(* IEC 61131-3 sources: daoli-st-library/DL_Process (part 53) *)

(* ---- FB_DL_StringCurrentMismatch.st ---- *)
(*
  FB_DL_StringCurrentMismatch  —  组串电流失配诊断与遮挡定位 / PV string current mismatch diagnostics and shading localisation
  分类 Category : DL_Process
  码位 Code     : 16#06_0_84
  版本 Version  : 1.0.0
  溯源 Source   : LGF Measurement 语义借鉴 · clean-room 实现，仅借分类/参数域/命名，未复制源码
  功能 Function : 1) 剔除无效/停机串后取中位基线（中位数抗单串遮挡污染，优于均值）；
                  2) 按失配率分级，失配率分母（基线）近零时自动切换为绝对差判据，防除零；
                  3) 输出最劣串物理串号（连续编址 1..16，越界钳位并置码）与失配掩码。
  边界 Boundary : ① 中位基线计算前剔除无效/停机串（电流 <= 0 或 NaN），有效样本 < 3 时不出诊断结论；
                  ② 失配率分母近零时改绝对差判据（防除零）；
                  ③ 遮挡定位输出按物理串号连续编址，越界下标钳位并置码；
                  ④ 结论态三行同向：基线值 → 最劣串号 → 失配标志。
  依赖 Depends  : None

  码表 Error codes（本件子码步进 16#10，避让邻件码位）:
    16#0002_0684 故障级：串数配置越界（nStringCount 不在 1..16）
    16#0002_0694 故障级：物理串号越界（枚举兜底路径，索引钳位后仍不可能命中）
    16#0002_06A4 信息级：有效样本不足 3 串，本轮不出诊断结论（不置 bError）
*)

TYPE E_DL_ScmPhase :
(
    eIdle    := 0,   // 空闲 / Idle
    eCollect := 10,  // 采样与剔除 / Sampling and rejection
    eDiagnose:= 20,  // 诊断计算 / Diagnostic computation
    eVerdict := 30,  // 结论输出 / Verdict output
    eFault   := 90   // 故障锁定 / Fault locked
);
END_TYPE

FUNCTION_BLOCK FB_DL_StringCurrentMismatch
VAR_INPUT
    bEnable       : BOOL;                         // 总使能，FALSE 回空闲 / Master enable
    bSample       : BOOL := TRUE;                 // 采样使能，TRUE 每拍纳入诊断 / Sampling enable
    bReset        : BOOL;                         // 复位，上升沿清故障 / Reset, clears fault
    nStringCount  : INT := 16;                    // 组串总数 [串]，域 1~16 / String count, 1..16
    afCurrentA    : ARRAY[1..16] OF REAL;         // 各串电流 [A]，域 > 0 为有效 / Per-string current [A]
    abStringValid : ARRAY[1..16] OF BOOL;         // 各串通讯/熔断有效标志 / Per-string valid flag
    fMismatchPct  : REAL := 10.0;                 // 失配率告警门限 [%]，域 0~100 / Mismatch rate alarm limit [%]
    fAbsFloorA    : REAL := 0.5;                  // 基线近零时的绝对差门限 [A]，域 > 0 / Absolute-difference limit [A]
    fBaselineEpsA : REAL := 0.1;                  // 基线近零判据容差 [A]，域 > 0 / Baseline near-zero tolerance [A]
    fMinSample    : INT := 3;                     // 最少有效样本数 [串]，常量 3 / Minimum valid sample count
END_VAR
VAR_OUTPUT
    fBaselineA    : REAL;                         // 中位基线电流 [A] / Median baseline current [A]
    nWorstIdx     : INT;                          // 最劣串物理串号 1..16，0 = 无 / Worst string number, 0 = none
    fWorstDevPct  : REAL;                         // 最劣串失配率 [%] / Worst string mismatch rate [%]
    fWorstDevA    : REAL;                         // 最劣串绝对偏差 [A] / Worst string absolute deviation [A]
    abMismatchMask : ARRAY[1..16] OF BOOL;        // 失配掩码 [开关]，索引 = 物理串号 / Mismatch mask per physical string
    nMismatchCount : INT;                         // 失配串数 [串] / Mismatched string count
    bMismatch     : BOOL;                         // 存在失配（保持型）/ Mismatch present, held
    bEnoughSample : BOOL;                         // 样本数满足结论条件 / Enough samples for a verdict
    bError        : BOOL;                         // 故障标志，与故障级码配对 / Fault flag paired with fault codes
    uErrorId      : UDINT;                        // 事件码，0 = 无事件 / Event code, 0 = none
    eStateOut     : E_DL_ScmPhase;                // 状态机当前态，段尾单点映射 / Phase mapped at tail
END_VAR
VAR
    _eState       : E_DL_ScmPhase := E_DL_ScmPhase.eIdle;  // 内部状态 / Internal state
    rtrReset      : R_TRIG;                       // 复位沿 / Reset edge
    nN            : INT;                          // 钳位后串数 [串] / Clamped string count
    nI            : INT;                          // 串循环下标 / String loop index
    nJ            : INT;                          // 排序内层下标 / Sort inner index
    nValid        : INT;                          // 有效串数 [串] / Valid string count
    nClampCode    : INT;                          // 下标钳位次数 [次] / Index clamping count
    afSort        : ARRAY[1..16] OF REAL;         // 有效电流排序缓存 [A] / Sorted valid currents [A]
    fTmp          : REAL;                         // 排序交换暂存 [A] / Sort swap buffer [A]
    fMedian       : REAL;                         // 中位基线暂存 [A] / Median baseline buffer [A]
    fDev          : REAL;                         // 单串偏差暂存 [A] / Single-string deviation [A]
    fRate         : REAL;                         // 单串失配率暂存 [%] / Single-string rate [%]
    fWorst        : REAL;                         // 最劣偏差累计 [A] / Worst deviation accumulator [A]
    bNearZero     : BOOL;                         // 基线近零标志 / Baseline near-zero flag
    uFault        : UDINT;                        // 锁存故障码 / Latched fault code
    uInfo         : UDINT;                        // 信息级码 / Information code
END_VAR
VAR CONSTANT
    DL_SCM_STRMAX : INT := 16;                    // 组串数组上界 [串] / String array upper bound
    DL_SCM_PCTMAX : REAL := 100.0;                // 失配率上限 [%] / Mismatch rate ceiling [%]
END_VAR

(* === 段 0 · 实例刷新（无条件周期调用）=== *)
rtrReset(CLK := bReset);                          // 每拍刷新复位沿

(* === 段 1 · 组态与索引闸 === *)
nN := nStringCount;                               // 串数取用前钳位
IF nN < 1 THEN
    nN := 1;                                      // 下限钳位
END_IF
IF nN > DL_SCM_STRMAX THEN
    nN := DL_SCM_STRMAX;                          // 上限钳位
END_IF
IF (nStringCount < 1) OR (nStringCount > DL_SCM_STRMAX) THEN
    uFault := 16#0002_0684;                       // 故障级：串数配置越界
END_IF
IF rtrReset.Q THEN
    uFault := 16#0000;                            // 复位沿清锁存
    bMismatch := FALSE;                           // 失配标志同步复位
    nWorstIdx := 0;                               // 最劣串号复位
END_IF

(* === 段 2 · 主状态机（ENUM + CASE，含 ELSE 兜底）=== *)
CASE _eState OF
E_DL_ScmPhase.eIdle :
    bEnoughSample := FALSE;                       // 空闲无结论
    uInfo := 16#0000;                             // 信息码清零
    IF uFault = 16#0002_0684 THEN
        _eState := E_DL_ScmPhase.eFault;          // 组态故障优先
    ELSIF bEnable AND bSample THEN
        _eState := E_DL_ScmPhase.eCollect;        // 本拍进入采样相
    END_IF

E_DL_ScmPhase.eCollect :
    nValid := 0;                                  // 有效串计数清零
    nClampCode := 0;                              // 钳位计数清零
    FOR nI := 1 TO DL_SCM_STRMAX DO
        IF nI <= nN THEN
            IF abStringValid[nI]
               AND (afCurrentA[nI] = afCurrentA[nI])              // NaN 自反判据
               AND (ABS(afCurrentA[nI]) < 1.0E30)                 // Inf 上限兜底
               AND (afCurrentA[nI] > 0.0) THEN                    // 停机串（<= 0）剔除
                nValid := nValid + 1;                             // 有效样本计数
                afSort[nValid] := afCurrentA[nI];                 // 收入排序缓存，nValid 已受 DL_SCM_STRMAX 约束
            END_IF
        END_IF
    END_FOR
    IF fMinSample < 3 THEN
        fMinSample := 3;                          // 最小样本数下限钳位（域 >= 3，防组态放宽到误判）
    END_IF
    bEnoughSample := (nValid >= fMinSample);      // 样本不足不出结论
    IF bEnoughSample THEN
        _eState := E_DL_ScmPhase.eDiagnose;       // 转诊断相
    ELSE
        uInfo := 16#0002_06A4;                    // 信息级：样本不足
        _eState := E_DL_ScmPhase.eVerdict;        // 仍走结论相，但结论为空
    END_IF

E_DL_ScmPhase.eDiagnose :
    FOR nI := 1 TO (nValid - 1) DO                // 插入排序求中位数
        FOR nJ := nI + 1 TO nValid DO
            IF afSort[nJ] < afSort[nI] THEN
                fTmp := afSort[nI];               // 交换暂存
                afSort[nI] := afSort[nJ];
                afSort[nJ] := fTmp;
            END_IF
        END_FOR
    END_FOR
    IF (nValid MOD 2) = 1 THEN
        fMedian := afSort[(nValid + 1) / 2];      // 奇数：取正中样本，下标受 nValid 约束
    ELSE
        fMedian := (afSort[nValid / 2] + afSort[(nValid / 2) + 1]) * 0.5;   // 偶数：取中两样本均值
    END_IF
    fBaselineA := fMedian;                        // 基线输出
    bNearZero := (ABS(fMedian) <= fBaselineEpsA); // 基线近零判据（防除零前置）
    nWorstIdx := 0;                               // 最劣串号先清零
    fWorst := -1.0;                               // 最劣偏差累计初值（负值确保首次必更新）
    fWorstDevPct := 0.0;                          // 最劣失配率初值
    fWorstDevA := 0.0;                            // 最劣绝对偏差初值
    nMismatchCount := 0;                          // 失配串计数清零
    FOR nI := 1 TO DL_SCM_STRMAX DO
        abMismatchMask[nI] := FALSE;              // 掩码逐串先清零
        IF nI <= nN THEN
            IF abStringValid[nI] AND (afCurrentA[nI] = afCurrentA[nI]) AND (afCurrentA[nI] > 0.0) THEN
                fDev := fMedian - afCurrentA[nI];                 // 偏差 = 基线 − 实测（正 = 偏低）
                IF bNearZero THEN
                    fRate := ABS(fDev);                               // 基线近零：改绝对差判据
                ELSE
                    fRate := ABS(fDev) / ABS(fMedian) * DL_SCM_PCTMAX;   // 分母已判非零
                END_IF
                IF fRate > DL_SCM_PCTMAX THEN
                    fRate := DL_SCM_PCTMAX;                       // 失配率饱和，防超界显示
                END_IF
                IF (bNearZero AND (ABS(fDev) > fAbsFloorA))
                   OR ((NOT bNearZero) AND (fRate >= fMismatchPct)) THEN
                    abMismatchMask[nI] := TRUE;                   // 该串判失配
                    nMismatchCount := nMismatchCount + 1;         // 失配计数累加
                END_IF
                IF fDev > fWorst THEN
                    fWorst := fDev;                               // 记录最劣偏差
                    IF (nI >= 1) AND (nI <= DL_SCM_STRMAX) THEN
                        nWorstIdx := nI;                          // 物理串号连续编址
                    ELSE
                        nWorstIdx := 0;                           // 越界下标钳位为 0
                        nClampCode := nClampCode + 1;             // 记录钳位事件
                    END_IF
                    fWorstDevPct := fRate;                        // 最劣串失配率
                    fWorstDevA := ABS(fDev);                      // 最劣串绝对偏差
                END_IF
            END_IF
        END_IF
    END_FOR
    bMismatch := (nMismatchCount > 0);            // 置位型结论：存在失配（段尾不清零）
    IF nClampCode > 0 THEN
        uFault := 16#0002_0694;                   // 故障级：物理串号越界已钳位
    END_IF
    _eState := E_DL_ScmPhase.eVerdict;            // 转结论相

E_DL_ScmPhase.eVerdict :
    IF NOT bEnoughSample THEN
        nWorstIdx := 0;                           // 样本不足：不给定位结论
        nMismatchCount := 0;                      // 失配计数归 0
        fWorstDevPct := 0.0;                      // 失配率归 0，避免误导
    END_IF
    IF (NOT bEnable) OR rtrReset.Q THEN
        _eState := E_DL_ScmPhase.eIdle;           // 失能/复位回空闲
    ELSIF bSample THEN
        _eState := E_DL_ScmPhase.eCollect;        // 连续采样：下一拍重新采集
    END_IF

E_DL_ScmPhase.eFault :
    bEnoughSample := FALSE;                       // 故障态不出结论
    nWorstIdx := 0;                               // 最劣串号 0
    IF uFault = 16#0000 THEN
        _eState := E_DL_ScmPhase.eIdle;           // 解锁后回空闲
    END_IF

ELSE
    _eState := E_DL_ScmPhase.eFault;              // 非法状态拦截
    uFault := 16#0002_0694;                       // 故障级：相 ID 越界（枚举兜底路径）
END_CASE

(* === 段 3 · 输出映射（三行同向：基线 → 最劣串号 → 失配标志）=== *)
IF NOT bEnoughSample THEN
    fBaselineA := fMedian;                        // 基线仍输出（诊断可读）
    bMismatch := nMismatchCount > 0;               // 失配标志与计数严格同源
END_IF
IF NOT bEnable THEN
    bMismatch := FALSE;                           // 失能强制清失配结论
    nWorstIdx := 0;                               // 最劣串号归 0
END_IF
bError := (uFault <> 16#0000);                    // 故障标志仅由故障级码置位（R45 配对）
IF bError THEN
    uErrorId := uFault;                           // 故障级优先上报
ELSE
    uErrorId := uInfo;                            // 否则上报信息级码
END_IF
eStateOut := _eState;                             // 输出枚举段尾单点映射（N2 规则）
END_FUNCTION_BLOCK

(* ---- FB_DL_StringElImageMap.st ---- *)
(*
  ==================================================================
  组件名 Component  : FB_DL_StringElImageMap
  分类   Category   : DL_Process
  版本   Version    : 1.0.1
  功能   Purpose    : EL 图像缺陷坐标归档与批次比对。逐条接收缺陷报告（坐标、面积、
                      类型），回钳后写入环窗归档（最新 64 条），并按批号累计本批
                      缺陷数、面积和 / 最大值 / 类型掩码；批号变化沿把当前批统计
                      转入「上批」快照并清零当前批，随后给出与上批的比对结论
                      （缺陷数与最大面积双向带容差比较）。
  溯源   Origin     : 缺陷坐标归档与批次间对比为通用视觉质量统计语义；本件为
                      clean-room 实现，仅借鉴来源分类与参数域组织（来源标签
                      roadmap-p2-elimage），道莅原创设计，未复制任何闭源代码行。
  平台   Platform   : 纯 IEC 61131-3（ARRAY / WORD / SHL / R_TRIG，无私有库）
  作者   Author     : 道莅代码库 · PLC 编程专家（R55）
  ------------------------------------------------------------------
  边界 Boundary     :
                      一 本件只做归档与统计比对，不做缺陷判定、不存图像（属主边界）；
                      二 坐标越出视野范围不归档，但计入越界计数并置信息级成因；
                      三 非有限坐标或面积不归档、不计数，出口数值保持上拍值；
                      四 环窗游标一律经回钳 1..64，写入顺序为「先算槽位、后写入」；
                      五 无全局变量、无外部变量声明、无物理地址寻址。
  输出契约 Output contract:
                      wTypeMask 位 i-1 对应缺陷类型 i（类型 1 得 bit0，类型 8 得 bit7）；
                      bComparePass 仅在无参照批（上批缺陷数为零）时恒为真，
                      有参照批时按「缺陷数」与「最大面积」双向带容差比较；
                      eCause 故障级成因与 bError 配对（R45），信息级永不置 bError。
  修订记录 Revision  :
    2026-11-20  v1.0.0  R55 首版（批 3 · 序号 12）
    2026-11-20  v1.0.1  R56 返修（7.4）：段 2 复位作用域补清 fLastXmm / fLastYmm /
                        fLastSizeMm2 / nLastType 四个最近缺陷出口，并补
                        _stCur.uBatchId 批号重同步，防复位后首条新批报告误判入旧批窗口。
  ==================================================================
*)

TYPE ST_DL_ElBatchStat :
STRUCT
    uBatchId  : UDINT := 0;      // 批号 [-] / batch identifier
    nCount    : INT := 0;        // 缺陷条数 [条] / defect count [piece]
    fSumSize  : REAL := 0.0;     // 面积累计 [平方毫米] / accumulated area [square millimetre]
    fMaxSize  : REAL := 0.0;     // 面积最大值 [平方毫米] / maximum area [square millimetre]
    wTypeMask : WORD := 16#0000; // 类型掩码 [-] / type mask
END_STRUCT
END_TYPE

TYPE E_DL_SeiCause :
(
    eNone       := 0,   // 无成因 / no cause
    eCfgIllegal := 1,   // 组态非法：视野范围或容差越域（故障级，与 bError 配对）/ illegal config, field bounds or tolerance out of domain
    eOutField   := 2,   // 缺陷坐标越出视野，未归档（信息级）/ the defect coordinate is outside the field and was not archived, informational
    eInputBad   := 3,   // 坐标或面积非有限，未归档（信息级）/ non-finite coordinate or area, not archived, informational
    eTypeBad    := 4    // 缺陷类型越域已回钳（信息级）/ the defect type was clamped, informational
);
END_TYPE

FUNCTION_BLOCK FB_DL_StringElImageMap
VAR_INPUT
    bEnable       : BOOL := TRUE;            // 使能，失能时不接收缺陷报告 [-] / enable, defect reports are not accepted when disabled
    bReset        : BOOL := FALSE;          // 复位上升沿清故障锁存与全部统计 [-] / reset rising edge clears the fault latch and all statistics
    bDefectValid  : BOOL := FALSE;           // 缺陷报告脉冲，上升沿归档一次 [-] / defect report pulse, archived once on the rising edge
    fPosXmm       : REAL := 0.0;             // 缺陷中心横坐标 [毫米] / defect centre abscissa [millimetre]
    fPosYmm       : REAL := 0.0;             // 缺陷中心纵坐标 [毫米] / defect centre ordinate [millimetre]
    fSizeMm2      : REAL := 0.0;             // 缺陷面积 [平方毫米] / defect area [square millimetre]
    nDefectType   : INT := 1;                // 缺陷类型 [类型号]，域 1..8 / defect type [type number], domain 1 to 8
    uBatchId      : UDINT := 0;              // 当前批号 [-] / current batch identifier
    fFieldXmm     : REAL := 1000.0;          // 视野横向范围 [毫米]，域 大于零 / field width [millimetre], domain above zero
    fFieldYmm     : REAL := 1000.0;          // 视野纵向范围 [毫米]，域 大于零 / field height [millimetre], domain above zero
    fTolPct       : REAL := 10.0;            // 批次比对容差 [百分比]，域 大于零 / batch comparison tolerance [percent], domain above zero
END_VAR
VAR_OUTPUT
    fLastXmm      : REAL := 0.0;             // 最近归档缺陷横坐标 [毫米] / abscissa of the last archived defect [millimetre]
    fLastYmm      : REAL := 0.0;             // 最近归档缺陷纵坐标 [毫米] / ordinate of the last archived defect [millimetre]
    fLastSizeMm2  : REAL := 0.0;             // 最近归档缺陷面积 [平方毫米] / area of the last archived defect [square millimetre]
    nLastType     : INT := 0;                // 最近归档缺陷类型 [类型号] / type of the last archived defect [type number]
    uArchiveCnt   : UDINT := 0;              // 累计归档缺陷数 [条] / total archived defects [piece]
    nBufCount     : INT := 0;                // 环窗当前条数 [条] / ring buffer occupancy [piece]
    nCurCount     : INT := 0;                // 当前批缺陷条数 [条] / current batch defect count [piece]
    fCurMaxMm2    : REAL := 0.0;             // 当前批最大缺陷面积 [平方毫米] / current batch maximum area [square millimetre]
    fCurMeanMm2   : REAL := 0.0;             // 当前批平均缺陷面积 [平方毫米] / current batch mean area [square millimetre]
    nPrevCount    : INT := 0;                // 上批缺陷条数 [条] / previous batch defect count [piece]
    fPrevMaxMm2   : REAL := 0.0;             // 上批最大缺陷面积 [平方毫米] / previous batch maximum area [square millimetre]
    fDeltaMaxPct  : REAL := 0.0;             // 最大面积相对变化 [百分比] / relative change of the maximum area [percent]
    bComparePass  : BOOL := FALSE;           // 批次比对通过 [-] / batch comparison passed
    wTypeMask     : WORD := 16#0000;         // 当前批缺陷类型掩码 [-] / current batch defect type mask
    nOutFieldCnt  : INT := 0;                // 越界缺陷计数（饱和到上限）[条] / out of field defect count, saturated [piece]
    eCause        : E_DL_SeiCause := E_DL_SeiCause.eNone; // 成因出口 [枚举] / cause outlet [enum]
    bError        : BOOL := FALSE;           // 故障锁存标志 [-] / fault latch flag
END_VAR
VAR
    rtDefect      : R_TRIG;                  // 缺陷报告沿检测，段 0 无条件刷新 / defect report edge detector, refreshed unconditionally in segment zero
    rtReset       : R_TRIG;                  // 复位沿检测，段 0 无条件刷新 / reset edge detector, refreshed unconditionally in segment zero
    _stCur        : ST_DL_ElBatchStat;       // 当前批统计 / current batch statistics
    _stPrev       : ST_DL_ElBatchStat;       // 上批统计快照 / previous batch statistics snapshot
    _eCause       : E_DL_SeiCause := E_DL_SeiCause.eNone;  // 信息级成因，每拍重算 / informational cause, recomputed every scan
    _eFaultCause  : E_DL_SeiCause := E_DL_SeiCause.eNone;  // 故障级成因，锁存至复位沿 / fault cause, latched until the reset edge
    _bFault       : BOOL := FALSE;           // 故障锁存位 [-] / fault latch bit
    _bInit        : BOOL := FALSE;           // 首扫初始化完成标志（R310）/ first scan initialisation flag
    _bCfgBad      : BOOL := FALSE;           // 组态非法判定 [-] / illegal configuration verdict
    _bInOk        : BOOL := FALSE;           // 本拍缺陷数据有限 [-] / this scan defect data finite
    _bInField     : BOOL := FALSE;           // 坐标在视野内 [-] / the coordinate is inside the field
    _bTypeClamped : BOOL := FALSE;           // 类型号被回钳 [-] / the type number was clamped
    _bBatchRoll   : BOOL := FALSE;           // 本拍发生批号变化 [-] / the batch identifier changed this scan
    _nTypeUse     : INT := 1;                // 钳定后的缺陷类型号 [类型号] / clamped defect type number
    _nIdx         : INT := 1;                // 环窗写入槽位（1 起，回钳 1..64）[槽号] / ring write slot, one-based, clamped one through sixty four
    _wTypeBit     : WORD := 16#0001;         // 类型位掩码，先移位后置位（R327）/ type bit mask, shift before setting
    _wMask        : WORD := 16#0000;         // 类型掩码工作字 / type mask working word
    _fMean        : REAL := 0.0;             // 均值工作值 [平方毫米] / mean working value [square millimetre]
    _fDeltaPct    : REAL := 0.0;             // 相对变化工作值 [百分比] / relative change working value [percent]
    _fPrevMaxB    : REAL := 0.0;             // 上批最大面积基线，用于除零闸 [平方毫米] / previous maximum baseline against division by zero [square millimetre]
    _fPrevCntB    : REAL := 0.0;             // 上批条数基线，用于除零闸 [条] / previous count baseline against division by zero [piece]
    _fCurMaxB     : REAL := 0.0;             // 当前批最大面积暂存 [平方毫米] / current maximum area held in a local [square millimetre]
    _fCurCntB     : REAL := 0.0;             // 当前批条数暂存 [条] / current count held in a local [piece]
    _afX          : ARRAY[1..64] OF REAL := [64(0.0)]; // 环窗横坐标归档 [毫米] / ring archive of abscissae [millimetre]
    _afY          : ARRAY[1..64] OF REAL := [64(0.0)]; // 环窗纵坐标归档 [毫米] / ring archive of ordinates [millimetre]
    _afSz         : ARRAY[1..64] OF REAL := [64(0.0)]; // 环窗面积归档 [平方毫米] / ring archive of areas [square millimetre]
    _anType       : ARRAY[1..64] OF INT := [64(0)];    // 环窗类型归档 [类型号] / ring archive of type numbers [type number]
END_VAR
VAR CONSTANT
    DL_SEI_BUF_MAX   : INT := 64;            // 环窗容量与槽位回钳上界 [条] / ring capacity and slot clamp upper bound
    DL_SEI_TYPE_MIN  : INT := 1;             // 缺陷类型下限 [类型号] / defect type floor [type number]
    DL_SEI_TYPE_MAX  : INT := 8;             // 缺陷类型上限（与掩码位宽一致）[类型号] / defect type ceiling matching the mask width [type number]
    DL_SEI_COUNT_MAX : INT := 30000;         // 单批缺陷条数上限，防溢出 [条] / per batch defect count ceiling against overflow [piece]
    DL_SEI_AREA_MAX  : REAL := 1.0E6;        // 缺陷面积量级上限 [平方毫米] / defect area magnitude ceiling [square millimetre]
    DL_SEI_TOL_MAX   : REAL := 500.0;        // 比对容差上限 [百分比] / comparison tolerance ceiling [percent]
    DL_SEI_MASK_NONE : WORD := 16#0000;      // 空掩码常量 [-] / empty mask constant
    DL_SEI_MASK_ONE  : WORD := 16#0001;      // 单位位常量 [-] / single bit constant
END_VAR

// 段 0｜沿检测无条件周期刷新（禁入分支）/ segment 0, unconditional refresh of the edge detectors, never inside a branch
rtDefect(CLK := bDefectValid); // 缺陷报告沿无条件刷新 / unconditional refresh of the defect edge
rtReset(CLK := bReset); // 复位沿无条件刷新 / unconditional refresh of the reset edge

// 段 1｜首扫初始化（R310）：统计与环窗从确定起点开始 / segment 1, first scan initialisation
IF NOT _bInit THEN // 首扫一拍 / the very first scan
    _bInit := TRUE; // 置首扫完成标志 / raise the first scan flag
    _bFault := FALSE; // 故障锁存清零 / clear the fault latch
    _eCause := E_DL_SeiCause.eNone; // 信息级成因清零 / clear the informational cause
    _eFaultCause := E_DL_SeiCause.eNone; // 故障级成因清零 / clear the fault cause
    _stCur.uBatchId := uBatchId; // 当前批号初始化 / initialise the current batch identifier
    _stPrev.uBatchId := 0; // 上批号清零 / clear the previous batch identifier
    _nIdx := 1; // 环窗槽位归位 / park the ring slot at one
END_IF

// 段 2｜复位沿作用域：清锁存 / 清统计 / 清环窗游标（归档数组保留，不作判据）/ segment 2, reset edge scope
IF rtReset.Q THEN // 复位沿 / reset edge
    _bFault := FALSE; // 作用域一：清故障锁存 / scope one, clear the fault latch
    _eFaultCause := E_DL_SeiCause.eNone; // 作用域一：清故障级成因 / scope one, clear the fault cause
    _stCur.nCount := 0; // 作用域二：清当前批条数 / scope two, clear the current batch count
    _stCur.fSumSize := 0.0; // 作用域二：清面积累计 / scope two, clear the accumulated area
    _stCur.fMaxSize := 0.0; // 作用域二：清面积最大值 / scope two, clear the maximum area
    _stCur.wTypeMask := DL_SEI_MASK_NONE; // 作用域二：清类型掩码 / scope two, clear the type mask
    _stPrev.nCount := 0; // 作用域二：清上批条数 / scope two, clear the previous count
    _stPrev.fSumSize := 0.0; // 作用域二：清上批面积累计 / scope two, clear the previous accumulated area
    _stPrev.fMaxSize := 0.0; // 作用域二：清上批最大面积 / scope two, clear the previous maximum area
    _stPrev.wTypeMask := DL_SEI_MASK_NONE; // 作用域二：清上批类型掩码 / scope two, clear the previous type mask
    fLastXmm := 0.0; // 作用域二：清最近横坐标出口（R56 返修补齐）/ scope two, clear the last abscissa outlet
    fLastYmm := 0.0; // 作用域二：清最近纵坐标出口（R56 返修补齐）/ scope two, clear the last ordinate outlet
    fLastSizeMm2 := 0.0; // 作用域二：清最近面积出口（R56 返修补齐）/ scope two, clear the last area outlet
    nLastType := 0; // 作用域二：清最近类型出口（R56 返修补齐）/ scope two, clear the last type outlet
    _stCur.uBatchId := uBatchId; // 作用域二：当前批号重同步，防复位后首条新批报告误判入旧批窗口（R56 返修补齐）/ scope two, resync the current batch identifier so the first report after a reset is not judged against a stale batch window
    _nIdx := 1; // 作用域三：清环窗槽位 / scope three, clear the ring slot cursor
    nBufCount := 0; // 作用域三：清环窗占用 / scope three, clear the ring occupancy
    uArchiveCnt := 0; // 作用域三：清累计归档数 / scope three, clear the total archived count
    nOutFieldCnt := 0; // 作用域三：清越界计数 / scope three, clear the out of field count
END_IF

// 段 3｜组态域闸（R151 全覆盖）：视野范围与比对容差 / segment 3, configuration domain gate over the field bounds and the tolerance
_bCfgBad := FALSE; // 组态非法预置假 / preset the illegal configuration verdict to false
IF (fFieldXmm <= 0.0) OR (fFieldXmm <> fFieldXmm) OR (fFieldXmm > DL_SEI_AREA_MAX) THEN // 横向视野越域 / field width out of domain
    _bCfgBad := TRUE; // 判非法 / mark illegal
END_IF
IF (fFieldYmm <= 0.0) OR (fFieldYmm <> fFieldYmm) OR (fFieldYmm > DL_SEI_AREA_MAX) THEN // 纵向视野越域 / field height out of domain
    _bCfgBad := TRUE; // 判非法 / mark illegal
END_IF
IF (fTolPct <= 0.0) OR (fTolPct > DL_SEI_TOL_MAX) OR (fTolPct <> fTolPct) THEN // 容量越域 / tolerance out of domain
    _bCfgBad := TRUE; // 判非法 / mark illegal
END_IF
IF _bCfgBad AND (NOT _bFault) THEN // 组态非法且未锁存 / illegal configuration and not yet latched
    _bFault := TRUE; // 置故障锁存 / raise the fault latch
    _eFaultCause := E_DL_SeiCause.eCfgIllegal; // 故障级成因 (R45 配对 bError) / fault grade cause paired with bError
END_IF

// 段 4｜批号变化：当前批统计转入上批快照，当前批清零 / segment 4, batch change moves the current statistics into the previous snapshot
_bBatchRoll := (uBatchId <> _stCur.uBatchId); // 批号变化判据 / batch change criterion
IF _bBatchRoll THEN // 批号变化 / the batch identifier changed
    _stPrev.uBatchId := _stCur.uBatchId; // 上批号继承 / the previous identifier inherits
    _stPrev.nCount := _stCur.nCount; // 上批条数快照 / snapshot the previous count
    _stPrev.fSumSize := _stCur.fSumSize; // 上批面积累计快照 / snapshot the previous accumulated area
    _stPrev.fMaxSize := _stCur.fMaxSize; // 上批最大面积快照 / snapshot the previous maximum area
    _stPrev.wTypeMask := _stCur.wTypeMask; // 上批类型掩码快照 / snapshot the previous type mask
    _stCur.uBatchId := uBatchId; // 当前批号推进 / advance the current identifier
    _stCur.nCount := 0; // 当前批条数清零 / clear the current count
    _stCur.fSumSize := 0.0; // 当前批面积累计清零 / clear the current accumulated area
    _stCur.fMaxSize := 0.0; // 当前批最大面积清零 / clear the current maximum area
    _stCur.wTypeMask := DL_SEI_MASK_NONE; // 当前批类型掩码清零 / clear the current type mask
END_IF

// 段 5｜缺陷归档：有限性闸 → 视野闸 → 类型回钳 → 环窗写入 → 统计累加 / segment 5, defect archiving chain
_eCause := E_DL_SeiCause.eNone; // 信息级成因每拍重算 / the informational cause is recomputed every scan
_bTypeClamped := FALSE; // 类型回钳标志预置假 / preset the type clamp flag to false
IF rtDefect.Q AND bEnable AND (NOT _bFault) THEN // 缺陷报告沿且使能无故障 / defect edge while enabled and unfaulted
    _bInOk := (fPosXmm = fPosXmm) AND ((fPosXmm - fPosXmm) = (fPosXmm - fPosXmm)) AND (fPosYmm = fPosYmm) AND ((fPosYmm - fPosYmm) = (fPosYmm - fPosYmm)) AND (fSizeMm2 = fSizeMm2) AND ((fSizeMm2 - fSizeMm2) = (fSizeMm2 - fSizeMm2)); // 坐标与面积有限性闸 / finiteness gate on coordinates and area
    _bInField := _bInOk AND (fPosXmm >= 0.0) AND (fPosXmm <= fFieldXmm) AND (fPosYmm >= 0.0) AND (fPosYmm <= fFieldYmm) AND (fSizeMm2 >= 0.0) AND (fSizeMm2 <= DL_SEI_AREA_MAX); // 视野与面积域闸 / field and area domain gate
    _nTypeUse := nDefectType; // 类型号直通 / the type number passes through
    IF _nTypeUse < DL_SEI_TYPE_MIN THEN // 下越界 / below the lower bound
        _nTypeUse := DL_SEI_TYPE_MIN; // 回钳到 1 / clamp to one
        _bTypeClamped := TRUE; // 置回钳标志 / raise the clamp flag
    ELSIF _nTypeUse > DL_SEI_TYPE_MAX THEN // 上越界 / above the upper bound
        _nTypeUse := DL_SEI_TYPE_MAX; // 回钳到 8 / clamp to eight
        _bTypeClamped := TRUE; // 置回钳标志 / raise the clamp flag
    END_IF
    IF NOT _bInOk THEN // 数据非有限 / data non-finite
        _eCause := E_DL_SeiCause.eInputBad; // 信息级成因：未归档 / informational cause, not archived
    ELSIF NOT _bInField THEN // 坐标或面积越域 / coordinate or area out of domain
        _eCause := E_DL_SeiCause.eOutField; // 信息级成因：越界未归档 / informational cause, out of field
        IF nOutFieldCnt < DL_SEI_COUNT_MAX THEN // 未达计数上限 / below the count ceiling
            nOutFieldCnt := nOutFieldCnt + 1; // 越界计数递增 / increment the out of field count
        END_IF
    ELSE
        // 段 5.1｜环窗写入：先算槽位再写入，槽位经回钳 1..64 / segment 5.1, ring write with the slot clamped one through sixty four
        _nIdx := _nIdx + 1; // 槽位前移 / advance the slot
        IF _nIdx > DL_SEI_BUF_MAX THEN // 越过上界 / past the upper bound
            _nIdx := 1; // 回钳到一号槽 / clamp back to slot one
        END_IF
        _afX[_nIdx] := fPosXmm; // 横坐标归档 / archive the abscissa
        _afY[_nIdx] := fPosYmm; // 纵坐标归档 / archive the ordinate
        _afSz[_nIdx] := fSizeMm2; // 面积归档 / archive the area
        _anType[_nIdx] := _nTypeUse; // 类型归档 / archive the type
        IF nBufCount < DL_SEI_BUF_MAX THEN // 环窗未满 / the ring is not yet full
            nBufCount := nBufCount + 1; // 占用递增 / increment the occupancy
        END_IF
        IF uArchiveCnt < 2000000000 THEN // 累计计数未达保护上限（常量在 DINT 可表范围内）/ the total count is below the guard ceiling, the constant fits in DINT
            uArchiveCnt := uArchiveCnt + 1; // 累计归档数递增 / increment the total archived count
        END_IF
        fLastXmm := fPosXmm; // 最近横坐标出口 / last abscissa outlet
        fLastYmm := fPosYmm; // 最近纵坐标出口 / last ordinate outlet
        fLastSizeMm2 := fSizeMm2; // 最近面积出口 / last area outlet
        nLastType := _nTypeUse; // 最近类型出口 / last type outlet
        // 段 5.2｜当前批统计累加 / segment 5.2, accumulate the current batch statistics
        IF _stCur.nCount < DL_SEI_COUNT_MAX THEN // 未达条数上限 / below the count ceiling
            _stCur.nCount := _stCur.nCount + 1; // 条数递增 / increment the count
        END_IF
        _stCur.fSumSize := _stCur.fSumSize + fSizeMm2; // 面积累计 / accumulate the area
        IF fSizeMm2 > _stCur.fMaxSize THEN // 面积最大值刷新 / refresh the maximum area
            _stCur.fMaxSize := fSizeMm2; // 更新最大值 / update the maximum
        END_IF
        _wTypeBit := SHL(DL_SEI_MASK_ONE, _nTypeUse - 1); // 类型位掩码，位移量 0..7 由类型回钳证明 / type bit mask, the shift zero through seven is proven by the type clamp
        _stCur.wTypeMask := _stCur.wTypeMask OR _wTypeBit; // 类型掩码置位 / set the type bit
        IF _bTypeClamped THEN // 类型被回钳 / the type was clamped
            _eCause := E_DL_SeiCause.eTypeBad; // 信息级成因 / informational cause
        END_IF
    END_IF
END_IF

// 段 6｜批次比对：双向带容差比较，参照批缺陷数为零时判通过 / segment 6, batch comparison with a two sided tolerance
_fCurMaxB := _stCur.fMaxSize; // 当前批最大面积 / the current maximum area
_fCurCntB := INT_TO_REAL(_stCur.nCount); // 当前批条数实数化 / the current count as a real
_fPrevMaxB := _stPrev.fMaxSize; // 上批最大面积 / the previous maximum area
_fPrevCntB := INT_TO_REAL(_stPrev.nCount); // 上批条数实数化 / the previous count as a real
IF (_fPrevMaxB > 0.0) THEN // 有参照批 / a reference batch exists
    _fDeltaPct := (_fCurMaxB - _fPrevMaxB) / _fPrevMaxB * 100.0; // 最大面积相对变化，除子已证大于零 / relative change of the maximum area, divisor proven positive
    bComparePass := (_fCurMaxB <= _fPrevMaxB * (1.0 + fTolPct / 100.0)) AND (_fPrevCntB <= 0.0 OR (_fCurCntB <= _fPrevCntB * (1.0 + fTolPct / 100.0))); // 数与面积双向比较，条数基线为零时只比面积 / the count and area are both compared, with a zero count baseline only the area is compared
ELSE // 无参照批 / no reference batch
    _fDeltaPct := 0.0; // 相对变化记零 / the relative change is zeroed
    bComparePass := TRUE; // 无参照按通过处理（不误判不合格）/ no reference passes so nothing is falsely rejected
END_IF

// 段 7｜统一出口 / segment 7, unified outlet
nCurCount := _stCur.nCount; // 当前批条数出口 / current count outlet
fCurMaxMm2 := _stCur.fMaxSize; // 当前批最大面积出口 / current maximum area outlet
_fMean := 0.0; // 均值预置零 / preset the mean to zero
IF _stCur.nCount > 0 THEN // 有条数才可算均值 / the mean needs at least one piece
    _fMean := _stCur.fSumSize / INT_TO_REAL(_stCur.nCount); // 均值，除子已证大于零 / mean, divisor proven positive
END_IF
fCurMeanMm2 := _fMean; // 当前批均值出口 / current mean outlet
nPrevCount := _stPrev.nCount; // 上批条数出口 / previous count outlet
fPrevMaxMm2 := _stPrev.fMaxSize; // 上批最大面积出口 / previous maximum area outlet
fDeltaMaxPct := _fDeltaPct; // 相对变化出口 / relative change outlet
wTypeMask := _stCur.wTypeMask; // 类型掩码出口 / type mask outlet
IF _bFault THEN // 故障锁存优先 / the fault latch takes priority
    eCause := _eFaultCause; // 故障级成因锁存回放 / the fault cause is replayed from the latch
ELSE
    eCause := _eCause; // 信息级成因直映 / the informational cause is mapped directly
END_IF
bError := _bFault; // 故障标志与锁存位同源 / the fault flag shares the latch source
END_FUNCTION_BLOCK

(* ---- FB_DL_StringerTrend.st ---- *)
(*
  FB_DL_StringerTrend  —  串焊机多通道焊接温度曲线在线监视 / Stringer multi-channel soldering temperature monitor
  分类 Category : DL_Process
  码位 Code     : 16#06_0_8E
  版本 Version  : 1.0.0
  溯源 Source   : LGF Measurement 语义借鉴 · clean-room 实现，仅借分类/参数域/命名，未复制源码
  功能 Function : 1) 逐通道焊接温度峰值窗判定（窗口均值 ± 带宽 → OK / 偏高 / 偏高三档）；
                  2) 首异常通道号输出 + 批次综合 bBatchOk；
                  3) 告警出口经 FB_DL_AlarmManager 分级（通道 i → 报警通道 i）。
  边界 Boundary : ① 通道数 < 2 不出统计结论（单点无峰谷可言，组态闸拒算）；
                  ② 任一通道实测无效（NaN/幅值越域）从统计剔除并在 abChanMask 标出；
                  ③ 链速为 0 时峰值窗不外推：保持上次窗并置 bHold；
                  ④ 分档边界按 R28 终审二式覆盖「正好整除」与「上限 + 1」两条向量（容差闭区间归属）；
                  ⑤ 输出三行同向：通道分档 → 首异常通道 → 批次结论。
  依赖 Depends  : FB_DL_SignalStatistics × 16（逐通道统计，每拍无条件调用）
                  FB_DL_AlarmManager × 1（分级告警出口，每拍无条件调用）

  码表 Error codes（本件子码步进 16#10，避让邻件码位）:
    16#0002_068E 故障级：组态非法（通道数 < 2 或 > 16 / 峰值带宽 <= 0 / 告警优先级表越界）
    16#0002_069E 故障级：相 ID 越界（枚举兜底路径）
    16#0002_06AE 信息级：链速为 0 峰值窗保持 / 有效通道不足 2 本拍不出结论（不置 bError）
*)

TYPE E_DL_StrBand :
(
    eOk     := 0,   // 峰值在窗内 / Peak in window
    eHigh   := 10,  // 峰值偏高 / Peak above window
    eLow    := 20,  // 峰值偏低 / Peak below window
    eFrozen := 30   // 通道无效冻结 / Channel frozen by invalid input
);
END_TYPE

TYPE E_DL_StrPhase :
(
    eIdle    := 0,  // 空闲 / Idle
    eWatch   := 10, // 在线监视 / Online monitoring
    eHold    := 20, // 链速为 0 窗保持 / Window held at zero chain speed
    eFault   := 90  // 组态故障锁定 / Configuration fault locked
);
END_TYPE

FUNCTION_BLOCK FB_DL_StringerTrend
VAR_INPUT
    bEnable       : BOOL;                           // 总使能，FALSE 回空闲 / Master enable
    bReset        : BOOL;                           // 复位，上升沿清组态故障 / Reset, clears configuration fault
    aTempC        : ARRAY[1..16] OF REAL;           // 各通道焊接温度 [°C] / Channel soldering temperature [degC]
    nChanCount    : INT := 12;                      // 通道数 [路]，2..16 / Channel count
    fChainSpd     : REAL := 40.0;                   // 链速 [mm/s]，0 = 停链 / Chain speed [mm/s]
    fPeakBandK    : REAL := 8.0;                    // 峰值窗半宽 [K]，域 > 0 / Peak window half width [K]
    fPeakBaseC    : REAL := 235.0;                  // 峰值窗中心基准 [°C] / Peak window center [degC]
    nStatWindow   : INT := 32;                      // 统计窗口长度 [样本] / Statistics window length [sample]
    uHoldScans    : UINT := 10;                     // 链速 0 保持确认拍数 [拍] / Zero-speed hold confirm scans
    fEps          : REAL := 1.0E-6;                 // 浮点判零容差 [1] / Floating zero tolerance
END_VAR
VAR_OUTPUT
    aeBand        : ARRAY[1..16] OF E_DL_StrBand;   // 逐通道峰值窗分档 / Per-channel band judgment
    nFirstAbnChan : INT;                            // 首异常通道号 1..16，0 = 无 / First abnormal channel
    bBatchOk      : BOOL;                           // 批次综合结论（全部有效通道在窗）/ Batch overall verdict
    bHold         : BOOL;                           // 链速为 0 窗保持标志 / Zero-speed window hold flag
    abChanMask    : ARRAY[1..16] OF BOOL;           // 通道无效掩码（TRUE = 剔除）/ Channel invalid mask
    bError        : BOOL;                           // 故障标志，与故障级码配对 / Fault flag
    uErrorId      : UDINT;                          // 事件码，0 = 无事件 / Event code
    eStateOut     : E_DL_StrPhase;                  // 状态机当前态，段尾单点映射 / Phase mapped at tail
END_VAR
VAR
    _eState       : E_DL_StrPhase := E_DL_StrPhase.eIdle;  // 内部状态 / Internal state
    afbStat       : ARRAY[1..16] OF FB_DL_SignalStatistics;  // 逐通道统计实例（无条件调用）/ Per-channel statistics
    fbAlm         : FB_DL_AlarmManager;             // 分级告警实例（无条件调用）/ Alarm manager instance
    rtrReset      : R_TRIG;                         // 复位沿 / Reset edge
    abAlmSrc      : ARRAY[0..15] OF BOOL;           // 告警源打包（通道 i-1）/ Alarm source packing
    auPrio        : ARRAY[0..15] OF USINT;          // 告警优先级表（警告级）/ Alarm priority table
    bCfgOk        : BOOL;                           // 组态合法标志 / Configuration valid
    bChanOk       : BOOL;                           // 单通道本拍有效 / Single channel valid this scan
    bWinOk        : BOOL;                           // 统计窗已就绪（bStatValid）/ Statistics window ready
    bOutWin       : BOOL;                           // 峰值越窗（电平）/ Peak out of window
    nValidCnt     : INT;                            // 有效通道计数 [路] / Valid channel count
    nI            : INT;                            // 遍历索引 / Loop index
    uZeroCnt      : UINT;                           // 链速 0 确认计数 [拍] / Zero-speed confirm counter
    uFault        : UDINT;                          // 锁存故障码 / Latched fault code
    uInfo         : UDINT;                          // 信息级码 / Information code
END_VAR
VAR CONSTANT
    DL_STR_CMAX   : INT := 16;                      // 通道数上限 [路] / Channel count upper bound
    DL_STR_INFMAX : REAL := 1.0E30;                 // 温度有限值幅值上限 [°C] / Temperature finite bound [degC]
END_VAR

(* === 段 0 · 实例刷新 === *)
rtrReset(CLK := bReset);                          // 每拍刷新复位沿

(* === 段 1 · 组态闸 === *)
bCfgOk := (nChanCount >= 2) AND (nChanCount <= DL_STR_CMAX)    // 通道数域闸（< 2 拒算）
          AND (fPeakBandK > fEps)                                // 峰值带宽正域
          AND (fPeakBaseC = fPeakBaseC) AND (ABS(fPeakBaseC) < DL_STR_INFMAX);  // 基准 NaN 自反 + 幅值
IF NOT bCfgOk THEN
    uFault := 16#0002_068E;                       // 故障级：组态非法
END_IF
IF rtrReset.Q AND bCfgOk THEN
    uFault := 16#0000;                            // 复位沿清锁存（解除路径可达）
END_IF
uInfo := 16#0000;                                 // 信息码每拍清零
FOR nI := 0 TO 15 DO
    auPrio[nI] := 2;                              // 全通道告警统一警告级
    abAlmSrc[nI] := FALSE;                        // 告警源本拍清零后重填
END_FOR

(* === 段 2 · 链速判定与逐通道统计（实例无条件调用）=== *)
IF ABS(fChainSpd) < fEps THEN
    uZeroCnt := uZeroCnt + UINT#1;                // 链速为 0：确认计数累加
    IF uZeroCnt >= uHoldScans THEN
        bHold := TRUE;                            // 连续 N 拍 0 速：窗保持
        uInfo := 16#0002_06AE;                    // 信息级：链速为 0 峰值窗保持
    END_IF
ELSE
    uZeroCnt := UINT#0;                           // 链速恢复：计数清零
    bHold := FALSE;                               // 保持解除（可达路径：链速恢复即解除）
END_IF
nValidCnt := 0;                                   // 有效通道计数清零
nFirstAbnChan := 0;                               // 首异常通道清零（本拍重算）
bBatchOk := TRUE;                                 // 批次结论先假设成立
FOR nI := 1 TO DL_STR_CMAX DO
    aeBand[nI] := E_DL_StrBand.eOk;               // 分档先取 OK（逐通道覆盖）
    IF nI <= nChanCount THEN
        bChanOk := (aTempC[nI] = aTempC[nI]) AND (ABS(aTempC[nI]) < DL_STR_INFMAX);  // NaN 自反 + 幅值闸
        abChanMask[nI] := NOT bChanOk;            // 无效掩码标出
        afbStat[nI](fIn := aTempC[nI],            // 统计实例无条件调用
                    bSample := bChanOk AND bEnable AND (NOT bHold),  // 无效/保持拍不采新样本
                    nWindow := nStatWindow,       // 窗口长度透传
                    bClear := rtrReset.Q);        // 复位沿清窗
        bWinOk := bChanOk AND afbStat[nI].bStatValid;   // 统计结论有效性（n >= 2）
        IF bChanOk THEN
            nValidCnt := nValidCnt + 1;           // 有效通道计数
        ELSE
            aeBand[nI] := E_DL_StrBand.eFrozen;   // 无效通道：冻结档
            bBatchOk := FALSE;                    // 存在无效通道批次不出 OK
        END_IF
        IF bWinOk THEN
            bOutWin := (afbStat[nI].fMax > fPeakBaseC + fPeakBandK + fEps)   // 峰值超上限（含容差）
                       OR (afbStat[nI].fMax < fPeakBaseC - fPeakBandK - fEps);  // 峰值低于下限
            IF bOutWin THEN
                IF afbStat[nI].fMax > fPeakBaseC THEN
                    aeBand[nI] := E_DL_StrBand.eHigh;   // 偏高档
                ELSE
                    aeBand[nI] := E_DL_StrBand.eLow;    // 偏低档
                END_IF
                bBatchOk := FALSE;                // 越窗通道拉低批次结论
                abAlmSrc[nI - 1] := TRUE;         // 告警源打包（0 基映射）
                IF nFirstAbnChan = 0 THEN
                    nFirstAbnChan := nI;          // 首异常通道记录
                END_IF
            END_IF
        ELSE
            IF bChanOk AND (nValidCnt >= 1) AND (nValidCnt < 2) THEN
                uInfo := 16#0002_06AE;            // 信息级：有效通道不足 2 本拍不出结论
            END_IF
            bBatchOk := FALSE;                    // 统计未就绪不出批次 OK
        END_IF
    ELSE
        abChanMask[nI] := TRUE;                   // 超出组态通道数：掩码标出
        aeBand[nI] := E_DL_StrBand.eFrozen;       // 冻结档
    END_IF
END_FOR

(* === 段 3 · 告警实例（无条件调用）=== *)
fbAlm(abAlarmActive := abAlmSrc,                  // 逐通道告警源
      auPriority := auPrio,                       // 统一警告级
      bAck := rtrReset.Q,                         // 复位沿确认首出
      bEnable := bEnable AND bCfgOk);             // 使能且组态合法

(* === 段 4 · 主状态机（ENUM + CASE，含 ELSE 兜底）=== *)
CASE _eState OF
E_DL_StrPhase.eIdle :
    IF uFault <> 16#0000 THEN
        _eState := E_DL_StrPhase.eFault;          // 故障优先
    ELSIF bEnable AND bCfgOk THEN
        _eState := E_DL_StrPhase.eWatch;          // 使能进监视相
    END_IF

E_DL_StrPhase.eWatch :
    IF (uFault <> 16#0000) OR (NOT bEnable) THEN
        _eState := E_DL_StrPhase.eFault;          // 故障/失能转出
    ELSIF bHold THEN
        _eState := E_DL_StrPhase.eHold;           // 链速 0 转窗保持相
    END_IF

E_DL_StrPhase.eHold :
    IF (uFault <> 16#0000) OR (NOT bEnable) THEN
        _eState := E_DL_StrPhase.eFault;          // 故障/失能转出
    ELSIF NOT bHold THEN
        _eState := E_DL_StrPhase.eWatch;          // 链速恢复回监视（解除路径可达）
    END_IF

E_DL_StrPhase.eFault :
    IF uFault = 16#0000 THEN
        _eState := E_DL_StrPhase.eIdle;           // 解锁回空闲
    END_IF

ELSE
    _eState := E_DL_StrPhase.eFault;              // 非法状态拦截
    uFault := 16#0002_069E;                       // 故障级：相 ID 越界
END_CASE

(* === 段 5 · 输出映射 === *)
bError := (uFault <> 16#0000);                    // 故障标志仅由故障级码置位（R45 配对）
IF bError THEN
    uErrorId := uFault;                           // 故障级优先上报
ELSE
    uErrorId := uInfo;                            // 否则上报信息级码
END_IF
eStateOut := _eState;                             // 输出枚举段尾单点映射（N2 规则）
END_FUNCTION_BLOCK

(* ---- FB_DL_StringIrrNormalize.st ---- *)
(*
  ==================================================================
  组件名 Component  : FB_DL_StringIrrNormalize
  分类   Category   : DL_Process
  版本   Version    : 1.0.0
  功能   Purpose    : 组串电流辐照归一化。把实测组串电流归一到参考辐照（默认
                      1000 瓦每平方米）与参考电池温度（默认 25 摄氏度）下的等效
                      电流：分母 = (G / Gref) × [1 + k × (T − Tref)]，
                      分子 = 实测电流；归一化电流 = 分子 / 分母。
                      用于不同辐照 / 温度工况下的组串横向比对与遮挡判别。
  溯源   Origin     : 辐照与温度归一为公开光伏工程口径；本件为 clean-room 实现，
                      仅借鉴来源分类与参数域组织（来源标签 roadmap-p2-string），
                      道莅原创设计，未复制任何闭源代码行。
  平台   Platform   : 纯 IEC 61131-3（REAL 运算，无私有库、无方言转换）
  作者   Author     : 道莅代码库 · PLC 编程专家（R55）
  ------------------------------------------------------------------
  边界 Boundary     :
                      一 本件只做归一化与有效性判定，不判组件故障、不做 MPPT（属主边界）；
                      二 辐照低于有效下限（默认 50 瓦每平方米）时不归一，出口保持上拍值；
                      三 分母（辐照相对量 × 温度因子）低于 1E-6 时不归一，出口保持上拍值；
                      四 温度补偿可按 bTempComp 关闭，关闭时温度因子恒为 1；
                      五 无全局变量、无外部变量声明、无物理地址寻址。
  输出契约 Output contract:
                      fINormA 仅在 bValid 为真的拍更新，其余拍保持上一次有效值
                      （首拍保持引脚初值 0），非有限值永不写入出口；
                      nHoldCnt 为连续无效拍计数（上限饱和），供上层判「长时间不可归一」；
                      eCause 故障级成因与 bError 配对（R45），信息级永不置 bError。
  修订记录 Revision  :
    2026-11-20  v1.0.0  R55 首版（批 2 · 序号 10）
  ==================================================================
*)

TYPE E_DL_SinCause :
(
    eNone       := 0,   // 无成因 / no cause
    eCfgIllegal := 1,   // 组态非法：参考辐照、温度系数或参考温度越域（故障级，与 bError 配对）/ illegal config, reference irradiance, temperature coefficient or reference temperature out of domain
    eIrrLow     := 2,   // 辐照低于有效下限，本拍不归一（信息级）/ irradiance below the effective floor, not normalised this scan, informational
    eInputBad   := 3,   // 输入非有限或分母不可用，本拍不归一（信息级）/ non-finite input or unusable denominator, not normalised this scan, informational
    eDenormBad  := 4    // 分母超量程，结果不可信（信息级）/ the denominator is out of range and the result is untrustworthy, informational
);
END_TYPE

FUNCTION_BLOCK FB_DL_StringIrrNormalize
VAR_INPUT
    bEnable      : BOOL := TRUE;             // 使能，失能时冻结出口保持末值 [-] / enable, the outlet freezes and holds its last value when disabled
    bReset       : BOOL := FALSE;           // 复位上升沿清故障锁存与保持计数 [-] / reset rising edge clears the fault latch and the hold counter
    fIrrWm2      : REAL := 0.0;              // 实测辐照 [瓦每平方米] / measured irradiance [watt per square metre]
    fIMeasA      : REAL := 0.0;              // 实测组串电流 [安培] / measured string current [ampere]
    fCellTempC   : REAL := 25.0;             // 实测电池温度 [摄氏度] / measured cell temperature [degree Celsius]
    fIrrRefWm2   : REAL := 1000.0;           // 参考辐照 [瓦每平方米]，域 大于零 / reference irradiance [watt per square metre], domain above zero
    fTempRefC    : REAL := 25.0;             // 参考电池温度 [摄氏度] / reference cell temperature [degree Celsius]
    fTempCoefPct : REAL := 0.35;             // 温度系数 [百分比每开尔文]，域 0..2 / temperature coefficient [percent per Kelvin], domain 0 to 2
    fIrrMinWm2   : REAL := 50.0;             // 有效辐照下限 [瓦每平方米]，域 大于零 / effective irradiance floor [watt per square metre], domain above zero
    bTempComp    : BOOL := TRUE;             // 真 = 做温度补偿，假 = 温度因子恒为 1 [-] / true applies temperature compensation, false keeps the factor at one
    nHoldMax     : INT := 600;               // 连续无效拍计数上限 [拍]，域 1..100000 / hold counter ceiling [scan], domain 1 to 100000
END_VAR
VAR_OUTPUT
    fINormA      : REAL := 0.0;              // 归一化组串电流 [安培] / normalised string current [ampere]
    fDenom       : REAL := 0.0;              // 归一化分母（辐照相对量 × 温度因子）[无量纲] / normalisation denominator, relative irradiance times the temperature factor [dimensionless]
    fIRelPct     : REAL := 0.0;              // 辐照相对量 [百分比] / relative irradiance [percent]
    fTFac        : REAL := 1.0;              // 温度因子 [无量纲] / temperature factor [dimensionless]
    bValid       : BOOL := FALSE;            // 本拍归一结果是否有效 [-] / this scan result valid flag
    nHoldCnt     : INT := 0;                 // 连续无效拍计数（饱和到上限）[拍] / consecutive invalid scan count, saturated at the ceiling
    eCause       : E_DL_SinCause := E_DL_SinCause.eNone; // 成因出口 [枚举] / cause outlet [enum]
    bError       : BOOL := FALSE;            // 故障锁存标志 [-] / fault latch flag
END_VAR
VAR
    rtReset      : R_TRIG;                   // 复位沿检测，段 0 无条件刷新 / reset edge detector, refreshed unconditionally in segment zero
    _eCause      : E_DL_SinCause := E_DL_SinCause.eNone;  // 信息级成因，每拍重算 / informational cause, recomputed every scan
    _eFaultCause : E_DL_SinCause := E_DL_SinCause.eNone;  // 故障级成因，锁存至复位沿 / fault cause, latched until the reset edge
    _bFault      : BOOL := FALSE;            // 故障锁存位 [-] / fault latch bit
    _bInit       : BOOL := FALSE;            // 首扫初始化完成标志（R310）/ first scan initialisation flag
    _bInOk       : BOOL := FALSE;            // 三项输入均有限 [-] / all three inputs finite
    _bCfgBad     : BOOL := FALSE;            // 组态非法判定 [-] / illegal configuration verdict
    _bDivOk      : BOOL := FALSE;            // 分母可用判定 [-] / denominator usable verdict
    _bValid      : BOOL := FALSE;            // 本拍有效内部位 [-] / internal validity bit of this scan
    _nHoldUse    : INT := 1;                 // 钳定后的保持计数上限 [拍] / clamped hold counter ceiling [scan]
    _nHoldCnt    : INT := 0;                 // 连续无效拍计数工作值 [拍] / consecutive invalid scan counter [scan]
    _fIrrRel     : REAL := 0.0;              // 辐照相对量工作值 [无量纲] / relative irradiance working value [dimensionless]
    _fTFac       : REAL := 1.0;              // 温度因子工作值 [无量纲] / temperature factor working value [dimensionless]
    _fDenom      : REAL := 0.0;              // 分母工作值 [无量纲] / denominator working value [dimensionless]
    _fNorm       : REAL := 0.0;              // 归一化结果工作值 [安培] / normalised result working value [ampere]
    _fNormHold   : REAL := 0.0;              // 归一化结果保持块 [安培] / normalised result holder [ampere]
END_VAR
VAR CONSTANT
    DL_SIN_DENOM_MIN : REAL := 1.0E-6;       // 分母下限，防除零 [无量纲] / denominator floor against division by zero [dimensionless]
    DL_SIN_DENOM_MAX : REAL := 1.0E3;        // 分母上限，防量纲错配放大 [无量纲] / denominator ceiling against a magnitude mismatch [dimensionless]
    DL_SIN_NORM_MAX  : REAL := 1.0E6;        // 归一化电流量级上限 [安培] / normalised current magnitude ceiling [ampere]
    DL_SIN_COEF_MIN  : REAL := 0.0;          // 温度系数下限 [百分比每开尔文] / temperature coefficient floor [percent per Kelvin]
    DL_SIN_COEF_MAX  : REAL := 2.0;          // 温度系数上限 [百分比每开尔文] / temperature coefficient ceiling [percent per Kelvin]
    DL_SIN_TREF_MIN  : REAL := -50.0;        // 参考温度下限 [摄氏度] / reference temperature floor [degree Celsius]
    DL_SIN_TREF_MAX  : REAL := 100.0;        // 参考温度上限 [摄氏度] / reference temperature ceiling [degree Celsius]
    DL_SIN_HOLD_MAX  : INT := 100000;        // 保持计数上限的钳定上限 [拍] / clamp ceiling of the hold counter [scan]
    DL_SIN_IRR_MAX   : REAL := 2000.0;       // 辐照量级上限，超此视为不可信 [瓦每平方米] / irradiance magnitude ceiling above which the value is untrustworthy [watt per square metre]
END_VAR

// 段 0｜复位沿无条件周期刷新（禁入分支）/ segment 0, unconditional refresh of the reset edge, never inside a branch
rtReset(CLK := bReset); // 复位沿无条件刷新 / unconditional refresh of the reset edge

// 段 1｜首扫初始化（R310）/ segment 1, first scan initialisation
IF NOT _bInit THEN // 首扫一拍 / the very first scan
    _bInit := TRUE; // 置首扫完成标志 / raise the first scan flag
    _bFault := FALSE; // 故障锁存清零 / clear the fault latch
    _eCause := E_DL_SinCause.eNone; // 信息级成因清零 / clear the informational cause
    _eFaultCause := E_DL_SinCause.eNone; // 故障级成因清零 / clear the fault cause
    _nHoldCnt := 0; // 保持计数清零 / clear the hold counter
    _fNormHold := 0.0; // 保持块清零 / clear the holder
END_IF

// 段 2｜复位沿作用域：清故障锁存 / 清保持计数（出口保持块不清，避免读数跳变）/ segment 2, reset edge scope
IF rtReset.Q THEN // 复位沿 / reset edge
    _bFault := FALSE; // 作用域一：清故障锁存 / scope one, clear the fault latch
    _eFaultCause := E_DL_SinCause.eNone; // 作用域一：清故障级成因 / scope one, clear the fault cause
    _nHoldCnt := 0; // 作用域二：清连续无效拍计数 / scope two, clear the consecutive invalid count
END_IF

// 段 3｜组态域闸（R151 全覆盖）：参考辐照、参考温度、温度系数、辐照下限、计数上限 / segment 3, configuration domain gate over every tuning pin
_bCfgBad := FALSE; // 组态非法预置假 / preset the illegal configuration verdict to false
IF (fIrrRefWm2 <= 0.0) OR (fIrrRefWm2 <> fIrrRefWm2) OR (fIrrRefWm2 > DL_SIN_IRR_MAX) THEN // 参考辐照越域 / reference irradiance out of domain
    _bCfgBad := TRUE; // 判非法 / mark illegal
END_IF
IF (fTempRefC < DL_SIN_TREF_MIN) OR (fTempRefC > DL_SIN_TREF_MAX) OR (fTempRefC <> fTempRefC) THEN // 参考温度越域 / reference temperature out of domain
    _bCfgBad := TRUE; // 判非法 / mark illegal
END_IF
IF (fTempCoefPct < DL_SIN_COEF_MIN) OR (fTempCoefPct > DL_SIN_COEF_MAX) OR (fTempCoefPct <> fTempCoefPct) THEN // 温度系数越域 / temperature coefficient out of domain
    _bCfgBad := TRUE; // 判非法 / mark illegal
END_IF
IF (fIrrMinWm2 <= 0.0) OR (fIrrMinWm2 <> fIrrMinWm2) OR (fIrrMinWm2 >= fIrrRefWm2) THEN // 辐照下限越域或与参考值矛盾 / irradiance floor out of domain or contradicting the reference
    _bCfgBad := TRUE; // 判非法 / mark illegal
END_IF
IF (nHoldMax < 1) OR (nHoldMax > DL_SIN_HOLD_MAX) THEN // 计数上限越域 / counter ceiling out of domain
    _bCfgBad := TRUE; // 判非法 / mark illegal
END_IF
IF _bCfgBad AND (NOT _bFault) THEN // 组态非法且未锁存 / illegal configuration and not yet latched
    _bFault := TRUE; // 置故障锁存 / raise the fault latch
    _eFaultCause := E_DL_SinCause.eCfgIllegal; // 故障级成因 (R45 配对 bError) / fault grade cause paired with bError
END_IF
_nHoldUse := nHoldMax; // 计数上限直通 / counter ceiling passes through
IF _nHoldUse < 1 THEN // 下越界 / below the lower bound
    _nHoldUse := 1; // 回钳到 1 / clamp to one
ELSIF _nHoldUse > DL_SIN_HOLD_MAX THEN // 上越界 / above the upper bound
    _nHoldUse := DL_SIN_HOLD_MAX; // 回钳到上限 / clamp to the ceiling
END_IF

// 段 4｜输入有限性闸：三项全有限才参与换算，任一非有限即保持上拍出口 / segment 4, input finiteness gate over all three measurements
_bInOk := (fIrrWm2 = fIrrWm2) AND ((fIrrWm2 - fIrrWm2) = (fIrrWm2 - fIrrWm2)) AND (fIMeasA = fIMeasA) AND ((fIMeasA - fIMeasA) = (fIMeasA - fIMeasA)) AND (fCellTempC = fCellTempC) AND ((fCellTempC - fCellTempC) = (fCellTempC - fCellTempC)); // 辐照、电流、温度三项有限性闸 / finiteness gate on irradiance, current and temperature
_eCause := E_DL_SinCause.eNone; // 信息级成因每拍重算 / the informational cause is recomputed every scan
_bValid := FALSE; // 本拍有效位预置假 / preset the validity bit to false
IF (NOT _bInOk) OR _bFault OR (NOT bEnable) THEN // 输入非有限、故障锁存或失能 / non-finite input, fault latched or disabled
    _eCause := E_DL_SinCause.eInputBad; // 信息级成因：不归一 / informational cause, not normalised
ELSE
    // 段 5｜温度因子：补偿关闭时恒为 1；补偿开启时按系数与温差展开 / segment 5, temperature factor computation
    _fTFac := 1.0; // 温度因子默认 1 / the temperature factor defaults to one
    IF bTempComp THEN // 补偿开启 / compensation enabled
        _fTFac := 1.0 + (fTempCoefPct / 100.0) * (fCellTempC - fTempRefC); // 因子，除子为常量 100.0 / factor with the constant divisor one hundred
        IF _fTFac < 0.05 THEN // 因子过小（极端温差外推）/ the factor is too small for a valid extrapolation
            _fTFac := 0.05; // 钳到下限，防分母趋零 / clamped to the floor against a vanishing denominator
        ELSIF _fTFac > 5.0 THEN // 因子过大 / the factor is too large
            _fTFac := 5.0; // 钳到上限 / clamped to the ceiling
        END_IF
    END_IF
    // 段 6｜辐照相对量与分母：辐照低于有效下限时不归一 / segment 6, relative irradiance and denominator
    _fIrrRel := fIrrWm2 / fIrrRefWm2; // 辐照相对量，除子已由域闸证明大于零 / relative irradiance, divisor proven positive by the domain gate
    _fDenom := _fIrrRel * _fTFac; // 分母 / denominator
    _bDivOk := (_fDenom >= DL_SIN_DENOM_MIN) AND (_fDenom <= DL_SIN_DENOM_MAX); // 分母在可用区间 / the denominator is inside the usable band
    IF (fIrrWm2 < fIrrMinWm2) OR (fIrrWm2 > DL_SIN_IRR_MAX) THEN // 辐照低于下限或超量程上限 / irradiance below the floor or above the magnitude ceiling
        _eCause := E_DL_SinCause.eIrrLow; // 信息级成因：辐照不可用 / informational cause, irradiance unusable
    ELSIF NOT _bDivOk THEN // 分母不可用 / the denominator is unusable
        _eCause := E_DL_SinCause.eDenormBad; // 信息级成因：分母超量程 / informational cause, denominator out of range
    ELSE
        _fNorm := fIMeasA / _fDenom; // 归一化电流，除子已证不小于 1E-6 / normalised current, divisor proven not below one micro unit
        IF (_fNorm <> _fNorm) OR ((_fNorm - _fNorm) <> (_fNorm - _fNorm)) OR (ABS(_fNorm) > DL_SIN_NORM_MAX) THEN // 结果非有限或超量级 / the result is non-finite or out of magnitude
            _eCause := E_DL_SinCause.eDenormBad; // 信息级成因：结果不可信 / informational cause, the result is untrustworthy
        ELSE
            _fNormHold := _fNorm; // 有效拍更新保持块（非有限不穿透出口）/ the holder is updated on a valid scan so nothing non-finite passes the outlet
            _bValid := TRUE; // 置本拍有效 / raise the this-scan validity
            _nHoldCnt := 0; // 有效拍清零连续无效计数 / clear the count on a valid scan
        END_IF
    END_IF
END_IF

// 段 7｜无效拍计数：饱和到钳定上限，防溢出翻转 / segment 7, invalid scan counting saturated at the clamped ceiling
IF (NOT _bValid) AND bEnable AND (NOT _bFault) THEN // 仅在使能且无故障时累计无效拍 / counting runs only while enabled and unfaulted
    IF _nHoldCnt < _nHoldUse THEN // 未达上限 / below the ceiling
        _nHoldCnt := _nHoldCnt + 1; // 计数递增 / increment the count
    END_IF
END_IF

// 段 8｜统一出口 / segment 8, unified outlet
fINormA := _fNormHold; // 归一化电流出口取保持块 / the normalised current outlet takes the holder
fDenom := _fDenom; // 分母出口 / denominator outlet
fIRelPct := _fIrrRel * 100.0; // 辐照相对量出口，乘常量 100.0 / relative irradiance outlet with the constant multiplier one hundred
fTFac := _fTFac; // 温度因子出口 / temperature factor outlet
bValid := _bValid AND (NOT _bFault); // 有效出口受故障锁存否决（挂状态量）/ the valid outlet is vetoed by the fault latch, a state quantity
nHoldCnt := _nHoldCnt; // 连续无效拍计数出口 / hold counter outlet
IF _bFault THEN // 故障锁存优先 / the fault latch takes priority
    eCause := _eFaultCause; // 故障级成因锁存回放 / the fault cause is replayed from the latch
ELSE
    eCause := _eCause; // 信息级成因直映 / the informational cause is mapped directly
END_IF
bError := _bFault; // 故障标志与锁存位同源 / the fault flag shares the latch source
END_FUNCTION_BLOCK

(* ---- FB_DL_StringIVTrace.st ---- *)
//==============================================================================
// 功能块：FB_DL_StringIVTrace ｜ 中文名称：组串 IV 曲线扫描与特征点提取
// 所属子库：DL_Process ｜ 版本：v1.0.0 ｜ 兼容：CODESYS V3.5+ / TwinCAT 3 / 汇川 InoProShop
// 功能描述：光伏组串 IV 扫描顺控——恒压步进扫描（fVCmdV 由 0 按步距
//           递增至扫描上限），每步等驻留窗并握手 bMeasReady 采样电压/
//           电流，特征点提取：Isc = 起始电压步电流（V 约为零）、Voc =
//           电流首次跌破开路阈值的步电压、Pmax/Vmp/Imp = 全程功率最大
//           步、FF = Pmax/(Voc·Isc)（填充因子）。Voc 捕获后可提前收扫
//           （曲线尾段无信息量）。测量步超时（tMeasTimeout 窗满仍未
//           就绪）→ 故障中止扫描。
// 开源溯源 (Origin)：道莅原创实现（参考 IEC 61829 光伏方阵 IV 特性现场测量 分类与参数域）
// 单位表：电压[V] / 电流[A] / 功率[W] / 步距[V] / 填充因子[无量纲] /
//         阈值电流[A] / 时间[ms]
// 错误码表：16#0005_01F0 信息级（扫描完成且 Voc/Isc/Pmax 全捕获，不置
//           bError）/ 16#0005_01F1 信息级（特征点降级：Voc 或 Isc 未
//           有效捕获，FF 置 0 照常输出，不置 bError）/ 16#0005_032D
//           故障级（组态非法：步距/上限/阈值 <= 0、时间窗 <= 0 或任一
//           输入非有限，置 bError）/ 16#0005_032E 故障级（测量步超时：
//           tMeasTimeout 窗满 bMeasReady 仍未就绪，扫描中止锁存，置
//           bError——该场景不可由 032D 的组态类判据观测，属运行握手
//           独立域）/ 16#0005_032F 故障级兜底（状态机落 ELSE，置
//           bError）
// 状态机：E_DL_IvTracePhase（四态：eIdle=0 / eSweep=10 / eDone=20 /
//           eFault=99），CASE 含 ELSE 兜底，ELSE 置 032F 并清扫描输出
// 边界行为：① 组态非法 → 故障态锁存，bReset 复位；② bAbort → 本拍
//           拒绝扫描推进、清命令电压，回空闲（中止不占相位，单拍标志
//           不外泄）；③ Voc 提前捕获 → 扫描立即收尾（曲线尾段无信息量，
//           缩短扫拍）；④ Voc/Isc 缺失 → FF 置 0 + 信息 01F1 降级照常
//           输出（除零防御，不置故障）；⑤ 未启动/故障态命令电压冻结
//           为 0 并 bValid := FALSE；⑥ eDone 等启动撤销回空闲（同拍
//           重启防抖，R39 范式）。
// 修订历史：v1.0.0 2026-11-17 首版（R24 派单 · ROADMAP P0 §228）
//==============================================================================

(*------------------------------------------------------------------------------
 * 枚举: E_DL_IvTracePhase（归属本功能块，同文件发布，全库唯一定义）
 * 含义: IV 扫描相位，每个成员在 CASE 中有且仅有一个标签。
 *-----------------------------------------------------------------------------*)
TYPE E_DL_IvTracePhase :
(
    eIdle   := 0,   // 空闲：等启动沿 / Idle, awaiting start edge
    eSweep  := 10,  // 扫描：步进采集中 / Sweep, stepping and sampling
    eDone   := 20,  // 完成：特征点锁存，等启动撤销 / Done, features latched, awaiting start drop
    eFault  := 99   // 故障：组态非法/测量超时/非法状态 / Fault, config, measurement timeout or illegal state
);
END_TYPE

FUNCTION_BLOCK FB_DL_StringIVTrace
VAR_INPUT
    bStart       : BOOL;                    // 启动请求 [—]，上升沿生效 / Start request, rising edge
    bAbort       : BOOL;                   // 中止请求 [—]，任意拍生效 / Abort request, effective on any scan
    bReset       : BOOL;                   // 故障复位 [—]，上升沿清故障态 / Fault reset, rising edge clears the fault state
    fMeasV       : LREAL;                  // 测量电压回读 [V] / Measured voltage feedback [V]
    fMeasI       : LREAL;                  // 测量电流回读 [A] / Measured current feedback [A]
    bMeasReady   : BOOL;                   // 测量就绪握手 [—]（每步采样条件） / Measurement ready handshake
    fVStepV      : LREAL := 0.5;           // 电压步距 [V]，须 > 0 / Voltage step [V], must be > 0
    fVMaxV       : LREAL := 50.0;          // 扫描电压上限 [V]，须 > 步距 / Sweep voltage ceiling [V], must exceed the step
    fIocThreshA  : LREAL := 0.002;         // 开路阈值电流 [A]，电流低于此判 Voc，须 > 0 / Open-circuit current threshold [A], must be > 0
    tStepDwell   : TIME  := T#50MS;        // 每步驻留窗 [ms]，须 > 0 / Per-step dwell window [ms]
    tMeasTimeout : TIME  := T#1S;          // 测量超时窗 [ms]，须 > 驻留窗（R100 配比） / Measurement timeout window [ms], must exceed the dwell
END_VAR
VAR_OUTPUT
    fVCmdV    : LREAL;                     // 扫描命令电压 [V]（给电子负载/扫频源） / Sweep command voltage [V]
    fVocV     : LREAL;                     // 开路电压特征点 [V]，未捕获为 0 / Open-circuit voltage feature [V], zero when not captured
    fIscA     : LREAL;                     // 短路电流特征点 [A]，未捕获为 0 / Short-circuit current feature [A], zero when not captured
    fPmaxW    : LREAL;                     // 最大功率点功率 [W] / Maximum power point [W]
    fVmpV     : LREAL;                     // 最大功率点电压 [V] / Maximum power point voltage [V]
    fImpA     : LREAL;                     // 最大功率点电流 [A] / Maximum power point current [A]
    fFillFactor : LREAL;                   // 填充因子 [无量纲]，Voc·Isc 无效时置 0 / Fill factor, zero when Voc or Isc invalid
    ePhase    : E_DL_IvTracePhase;         // 扫描相位 [—] / Sweep phase
    bTraceDone: BOOL;                      // 扫描完成 [—]（完成态电平） / Trace done, completion level
    eErr      : UDINT;                     // 错误码，0 = 无错，码位 16#0005_01F0 起信息级、16#0005_032D 起故障级（分带见错误码表） / Error code, 0 = no error, band info/fault per the code table
    bError    : BOOL;                      // 故障级标志，仅故障级错误置位 / Fault-class flag, set only on fault-level codes
    bValid    : BOOL;                      // 输出可用标志 / Outputs usable flag
END_VAR
VAR
    fbDwell   : TON;                       // 每步驻留计时（每拍无条件刷新）[ms] / Dwell timer, refreshed unconditionally
    fbMeasTo  : TON;                       // 测量超时计时（每拍无条件刷新）[ms] / Measurement timeout timer, refreshed unconditionally
    fbStart   : R_TRIG;                    // 启动沿检测（待机/故障分支同样无条件刷新） / Start edge detector, refreshed unconditionally
    _ePhase   : E_DL_IvTracePhase := E_DL_IvTracePhase.eIdle; // 当前相位 / Current phase
    _bCfgBad  : BOOL;                      // 组态非法锁存 / Illegal config latch
    _fVSweep  : LREAL;                     // 当前扫描电压 [V] / Current sweep voltage [V]
    _fVocCap  : LREAL;                     // Voc 捕获暂存 [V] / Voc capture staging [V]
    _fIscCap  : LREAL;                     // Isc 捕获暂存 [A] / Isc capture staging [A]
    _bVocOk   : BOOL;                      // Voc 捕获有效标志 / Voc captured flag
    _bIscOk   : BOOL;                      // Isc 捕获有效标志 / Isc captured flag
    _bInfoFull: BOOL;                      // 全捕获信息当拍标志 / Full-capture info flag of this scan
    _bInfoDeg : BOOL;                      // 降级信息当拍标志 / Degraded info flag of this scan
    _bIllegal : BOOL;                      // 非法状态标志 / Illegal state flag
    _bInit    : BOOL := FALSE;             // 首扫标志，初值 FALSE 取非判定 / First-scan flag, tested negated
END_VAR
VAR CONSTANT
    DL_IVT_INF    : LREAL := 1.7976931348623157E308; // LREAL 幅值上限 / LREAL magnitude ceiling
    DL_IVT_EPS    : LREAL := 1.0E-6;        // 浮点判零容差 [混合] / Float zero tolerance
    DL_IVT_ZERO   : LREAL := 0.0;           // 零值常量，避免裸字面量 [混合] / Zero constant, avoids a bare literal
    DL_IVT_FF_MIN : LREAL := 0.0;           // 填充因子下限 [无量纲] / Fill factor floor
    DL_IVT_FF_MAX : LREAL := 1.0;           // 填充因子上限 [无量纲] / Fill factor ceiling
END_VAR

(*------------------------------------------------------------------------------
 * 段 1｜每拍预置：命令电压安全侧清零，特征输出每拍重算，单拍标志预清零
 *      Command voltage cleared fail-safe, features recomputed, flags pre-cleared
 *-----------------------------------------------------------------------------*)
fVCmdV   := DL_IVT_ZERO;                 // 命令电压先清（安全侧；扫描态在段 3 重置） / Command voltage cleared first
fVocV    := DL_IVT_ZERO;                 // 特征出口每拍重算 / Feature outlets recomputed
fIscA    := DL_IVT_ZERO;                 // 特征出口每拍重算 / Feature outlets recomputed
fPmaxW   := DL_IVT_ZERO;                 // 特征出口每拍重算 / Feature outlets recomputed
fVmpV    := DL_IVT_ZERO;                 // 特征出口每拍重算 / Feature outlets recomputed
fImpA    := DL_IVT_ZERO;                 // 特征出口每拍重算 / Feature outlets recomputed
fFillFactor := DL_IVT_ZERO;              // 填充因子每拍重算 / Fill factor recomputed
eErr   := 16#0000_0000;                  // 错误码每拍重算 / Error code recomputed
bError := FALSE;                         // 故障标志每拍重算 / Fault flag recomputed
bValid := FALSE;                         // 可用标志每拍重算 / Usable flag recomputed
_bInfoFull := FALSE;                     // 全捕获信息预清零 / Full-capture info pre-cleared
_bInfoDeg  := FALSE;                     // 降级信息预清零 / Degraded info pre-cleared
_bIllegal  := FALSE;                     // 非法状态预清零 / Illegal flag pre-cleared

(*------------------------------------------------------------------------------
 * 段 2｜首扫初始化
 *      First-scan initialisation
 *-----------------------------------------------------------------------------*)
IF NOT _bInit THEN
    _ePhase  := E_DL_IvTracePhase.eIdle; // 相位空闲起步 / Phase starts idle
    _bCfgBad := FALSE;                   // 组态锁存清零 / Config latch cleared
    _fVSweep := DL_IVT_ZERO;             // 扫描电压从零起步 / Sweep voltage starts at zero
    _bInit   := TRUE;                    // 首扫只做一次 / The first scan runs once
END_IF

(*------------------------------------------------------------------------------
 * 段 3｜组态防御闸 + 沿检测无条件刷新（R40）
 *      Config gates and unconditional edge/timer refresh
 *-----------------------------------------------------------------------------*)
fbStart(CLK := bStart);                  // 启动沿检测 / Start edge detection
IF (fVStepV <> fVStepV) OR (ABS(fVStepV) > DL_IVT_INF)
   OR (fVMaxV <> fVMaxV) OR (ABS(fVMaxV) > DL_IVT_INF)
   OR (fIocThreshA <> fIocThreshA) OR (ABS(fIocThreshA) > DL_IVT_INF)
   OR (fMeasV <> fMeasV) OR (ABS(fMeasV) > DL_IVT_INF)
   OR (fMeasI <> fMeasI) OR (ABS(fMeasI) > DL_IVT_INF) THEN
    _bCfgBad := TRUE;                    // 非有限归组态非法锁存 / Non-finite folded into the config latch
END_IF
IF (NOT _bCfgBad) AND ((fVStepV <= DL_IVT_EPS) OR (fVMaxV <= fVStepV)
   OR (fIocThreshA <= DL_IVT_EPS) OR (tStepDwell <= T#0MS)
   OR (tMeasTimeout <= tStepDwell)) THEN
    _bCfgBad := TRUE;                    // 步距/上限/阈值/时间窗非法锁存（含 R100 配比：超时窗 > 驻留窗） / Step, ceiling, threshold and window domains latched
END_IF

(*------------------------------------------------------------------------------
 * 段 4｜双计时无条件刷新（R40：CASE 之外每拍必调）
 *      Two timers refreshed unconditionally per R40
 *-----------------------------------------------------------------------------*)
fbDwell(IN := (_ePhase = E_DL_IvTracePhase.eSweep) AND (NOT bAbort), PT := tStepDwell); // 步驻留窗 / Step dwell window
fbMeasTo(IN := (_ePhase = E_DL_IvTracePhase.eSweep) AND (NOT bAbort)
              AND (NOT bMeasReady), PT := tMeasTimeout); // 测量超时窗 / Measurement timeout window

(*------------------------------------------------------------------------------
 * 段 5｜相位机（CASE 含 ELSE 兜底；状态改写只出现在分支判据内，R39）
 *      Phase machine with ELSE fallback
 *-----------------------------------------------------------------------------*)
CASE _ePhase OF

    E_DL_IvTracePhase.eIdle:               // 空闲：启动沿且组态合法进扫描
        IF fbStart.Q AND (NOT _bCfgBad) THEN
            _fVSweep := DL_IVT_ZERO;       // 扫描电压归零起步 / Sweep voltage reset to zero
            _bVocOk  := FALSE;             // 捕获标志复位 / Capture flags reset
            _bIscOk  := FALSE;             // 捕获标志复位 / Capture flags reset
            _ePhase  := E_DL_IvTracePhase.eSweep; // 进扫描 / To sweep
        ELSIF fbStart.Q AND _bCfgBad THEN
            _ePhase := E_DL_IvTracePhase.eFault; // 组态非法进故障 / Illegal config to fault
        END_IF

    E_DL_IvTracePhase.eSweep:              // 扫描：采样、判 Voc、步进、收尾
        IF _bCfgBad OR bAbort THEN
            fVCmdV := DL_IVT_ZERO;         // 中止拍拒绝推进并清命令（拍 N 进入行为） / Abort scan rejects progress and clears the command
            _ePhase := E_DL_IvTracePhase.eIdle; // 拍 N+1 转出：回空闲（中止不占相位） / Back to idle, abort holds no phase
        ELSIF fbMeasTo.Q THEN
            _ePhase := E_DL_IvTracePhase.eFault; // 测量超时进故障 / Measurement timeout to fault
        ELSIF fbDwell.Q AND bMeasReady THEN
            IF (NOT _bIscOk) AND (_fVSweep <= fVStepV) THEN
                _fIscCap := fMeasI;        // Isc：起始电压步电流（V 约为零） / Isc from the first near-zero step
                _bIscOk  := TRUE;          // Isc 捕获有效 / Isc captured
            END_IF
            IF (NOT _bVocOk) AND (fMeasI < fIocThreshA) THEN
                _fVocCap := fMeasV;        // Voc：电流首次跌破开路阈值步电压 / Voc at the first sub-threshold step
                _bVocOk  := TRUE;          // Voc 捕获有效 / Voc captured
            END_IF
            IF (fMeasV * fMeasI) > fPmaxW THEN
                fPmaxW := fMeasV * fMeasI; // 最大功率点功率 [W] / Maximum power [W]
                fVmpV  := fMeasV;          // 最大功率点电压 [V] / MPP voltage
                fImpA  := fMeasI;          // 最大功率点电流 [A] / MPP current
            END_IF
            IF _bVocOk OR (_fVSweep + fVStepV > fVMaxV) THEN
                _ePhase := E_DL_IvTracePhase.eDone; // Voc 已捕获或达上限：收扫 / Voc captured or ceiling reached, close the sweep
            ELSE
                _fVSweep := _fVSweep + fVStepV; // 步进推进 / Step advance
            END_IF
        END_IF

    E_DL_IvTracePhase.eDone:               // 完成：等启动撤销回空闲（同拍重启防抖）
        IF NOT bStart THEN
            _ePhase := E_DL_IvTracePhase.eIdle; // 回空闲 / Back to idle
        END_IF

    E_DL_IvTracePhase.eFault:              // 故障：复位沿且组态恢复回空闲
        IF bReset AND (NOT _bCfgBad) THEN
            _ePhase := E_DL_IvTracePhase.eIdle; // 回空闲 / Back to idle
        END_IF

    ELSE                                   // 非法状态兜底（R21：CASE 必带 ELSE）
        _bIllegal := TRUE;                 // 标记非法状态 / Flag the illegal state
        fVCmdV := DL_IVT_ZERO;             // 命令电压清零（安全侧） / Command cleared, safe side
        _ePhase := E_DL_IvTracePhase.eFault; // 回故障态 / Back to fault
END_CASE

(*------------------------------------------------------------------------------
 * 段 6｜扫描命令出口与特征点换算（除零防御 + 填充因子钳域）
 *      Command outlet and feature scaling with divide guards
 *-----------------------------------------------------------------------------*)
IF _ePhase = E_DL_IvTracePhase.eSweep THEN
    fVCmdV := _fVSweep;                    // 扫描态命令电压 = 当前扫描点 / Sweep command equals the current point
END_IF
IF _bVocOk THEN
    fVocV := _fVocCap;                     // Voc 出口 / Voc outlet
END_IF
IF _bIscOk THEN
    fIscA := _fIscCap;                     // Isc 出口 / Isc outlet
END_IF
IF _bVocOk AND _bIscOk THEN
    IF ABS(_fVocCap * _fIscCap) > DL_IVT_EPS THEN
        fFillFactor := MIN(MAX(fPmaxW / (_fVocCap * _fIscCap), DL_IVT_FF_MIN), DL_IVT_FF_MAX); // 填充因子 [无量纲]，分母已闸且钳域 / Fill factor, denominator gated and clamped
    END_IF
    IF _ePhase = E_DL_IvTracePhase.eDone THEN
        _bInfoFull := TRUE;                // 全捕获完成（信息级） / Full capture done, info
    END_IF
ELSIF _ePhase = E_DL_IvTracePhase.eDone THEN
    _bInfoDeg := TRUE;                     // 特征点降级：Voc 或 Isc 未捕获，FF 置 0（信息级） / Degraded features, FF zero, info
END_IF

(*------------------------------------------------------------------------------
 * 段 7｜码位出口与放行（故障级码 3 行内置 bError，R45/R101 配对）
 *      Code outlet and release, fault codes paired with bError
 *-----------------------------------------------------------------------------*)
IF _bIllegal THEN
    eErr   := 16#0005_032F;                // 故障级：状态机兜底 / Fault: state machine fallback
    bError := TRUE;                        // 置故障标志 / Raise the fault flag
ELSIF _bCfgBad THEN
    eErr   := 16#0005_032D;                // 故障级：组态非法（触发前或扫描中漂移同域） / Fault: illegal configuration, drift folded
    bError := TRUE;                        // 置故障标志 / Raise the fault flag
ELSIF _ePhase = E_DL_IvTracePhase.eFault THEN
    eErr   := 16#0005_032E;                // 故障级：测量步超时（组态恢复后落此域即超时） / Fault: measurement timeout
    bError := TRUE;                        // 置故障标志 / Raise the fault flag
ELSIF _bInfoDeg THEN
    eErr := 16#0005_01F1;                  // 信息级：特征点降级 / Info: degraded features
ELSIF _bInfoFull THEN
    eErr := 16#0005_01F0;                  // 信息级：扫描完成全捕获 / Info: sweep done, full capture
END_IF

bTraceDone := (_ePhase = E_DL_IvTracePhase.eDone); // 完成电平挂状态量（R99） / Done level bound to the state
bValid := (NOT bError) AND (_ePhase = E_DL_IvTracePhase.eDone); // 仅完成态放行 / Usable only in the done phase
ePhase := _ePhase;                       // 相位出口 / Phase outlet
END_FUNCTION_BLOCK

(* ---- FB_DL_StringSolderQuality.st ---- *)
(*
  FB_DL_StringSolderQuality  —  串焊焊接质量在线判据 / String soldering quality online criteria
  分类 Category : DL_Process
  码位 Code     : 16#06_0_B4
  版本 Version  : 1.0.0
  来源 Source   : t2-1-lgf-technology — IEC 61131-3 标准语义的道莅防御性实现
  溯源 Origin   : clean-room 实现，光伏串焊温度曲线公开工艺语义借鉴，未复制任何源码行（RESUME 承接 R36 §4 #19 规格）
                  （统计出口语义对齐 FB_DL_SignalStatistics；告警出口对齐 FB_DL_AlarmManager，均不实例化）
  功能 Function : 1) 逐通道三判据：峰值窗（fPeakMinC..fPeakMaxC）、升温斜率窗、保温时长窗，越窗记 abPeakViolate/abSlopeViolate
                     （保温越窗并入 abPeakViolate 位段，头注释声明）并聚合 nNgChannelMask（SHL 显式位号）；
                  2) 拉力抽检仅对抽中通道（abPullSampled）生效，抽检不合格整批 bLotReject；
                  3) 曲线 NG 通道与抽检通道双判据独立记账，不互相掩盖。
  边界 Boundary : ① 通道数 nChannelCount = 0 或超 32 判组态错返回；
                  ② 位掩码只在 nChannelCount <= 32 时生成（超 32 判组态错，禁静默截断，规格强制）；
                  ③ fSlopeMaxCs <= fSlopeMinCs / fPeakMaxC <= fPeakMinC 判组态错；
                  ④ 信号非有限（NaN 用 x<>x 自反）通道按 NG 记（安全侧）并置信息码；
                  ⑤ 整数位段赋值用 SHL 显式位号，禁魔法掩码（规格强制）；
                  ⑥ 本件无状态机 ENUM/CASE（批量判据件），判据每调用重算，无锁存码。
  依赖 Depends  : 仅 Standard.library（SHL/AND_MASK）；语义对齐 FB_DL_SignalStatistics / FB_DL_AlarmManager（已注册，不实例化）
  码表 Error codes（本件格 06_0_B4，子码步进 +0x100）:
    16#0006_01B4 信息级：拉力抽检不合格，整批判废
    16#0006_02B4 故障级：组态非法（通道数越域 / 峰值窗倒置 / 斜率窗倒置 / 时长窗倒置）
    16#0006_03B4 信息级：存在曲线越窗通道（nNgChannelMask <> 0）
    16#0006_04B4 信息级：存在非有限信号通道，按 NG 记（安全侧）

  修订历史 Revision :
    2026-11-18  v1.0.0  R38 首版
*)

FUNCTION_BLOCK FB_DL_StringSolderQuality
VAR_INPUT
    afPeakC       : ARRAY[0..31] OF REAL;   // 各通道峰值温度 [°C] / Per-channel peak temperature
    afSlopeCs     : ARRAY[0..31] OF REAL;   // 各通道升温斜率 [°C/s] / Per-channel ramp slope
    afHoldMs      : ARRAY[0..31] OF REAL;   // 各通道保温时长 [ms] / Per-channel hold duration
    abPullSampled : ARRAY[0..31] OF BOOL;   // 拉力抽中通道表 / Pull-test sampled channels
    afPullN       : ARRAY[0..31] OF REAL;   // 抽检拉力值 [N] / Pull test force
    nChannelCount : INT;                    // 有效通道数 [路]，域 1..32 / Valid channel count
    fPeakMinC     : REAL := 220.0;          // 峰值窗下限 [°C] / Peak window floor
    fPeakMaxC     : REAL := 260.0;          // 峰值窗上限 [°C] / Peak window ceiling
    fSlopeMinCs   : REAL := 2.0;            // 斜率窗下限 [°C/s] / Slope window floor
    fSlopeMaxCs   : REAL := 10.0;           // 斜率窗上限 [°C/s] / Slope window ceiling
    fHoldMinMs    : REAL := 800.0;          // 保温时长窗下限 [ms] / Hold window floor
    fHoldMaxMs    : REAL := 3000.0;         // 保温时长窗上限 [ms] / Hold window ceiling
    fPullMinN     : REAL := 1.5;            // 拉力抽检下限 [N] / Pull test force floor
END_VAR
VAR_OUTPUT
    abChannelOk    : ARRAY[0..31] OF BOOL;  // 逐通道合格 / Per-channel verdict
    abPeakViolate  : ARRAY[0..31] OF BOOL;  // 逐通道峰值越窗（含保温越窗并入位段）/ Per-channel peak violation
    abSlopeViolate : ARRAY[0..31] OF BOOL;  // 逐通道斜率越窗 / Per-channel slope violation
    nNgChannelMask : DWORD;                 // NG 通道位掩码（<= 32 路才生成）/ NG channel bit mask
    bLotReject     : BOOL;                  // 整批判废 / Lot reject verdict
    nErrId         : UDINT;                 // 事件码，0 = 无事件 / Event code
END_VAR
VAR
    _nK        : INT;                       // 通道循环计数 / Channel loop counter
    _bFin      : BOOL;                      // 非有限筛查标志 / Non-finite screening flag
    _bPullFail : BOOL;                      // 拉力抽检失败聚合（独立记账）/ Pull failure aggregate
    _bAnyNg    : BOOL;                      // 任一通道 NG 聚合 / Any channel NG aggregate
    _bCfgBad   : BOOL;                      // 组态非法聚合 / Configuration invalid aggregate
    _uInfo     : UDINT;                     // 信息码，每拍重算 / Info code
END_VAR
VAR CONSTANT
    nMaxCh : INT := 32;           // 数组上界 = 掩码位宽 [路] / Array bound = mask width
END_VAR

(* —— 段 1：单拍量预清零（判据件每调用重算，无锁存量，R187①） —— *)
_uInfo := 16#0000_0000;              // 信息码每拍重算
nNgChannelMask := 0;                 // 掩码缺省 0
bLotReject := FALSE;                 // 判废缺省 FALSE
_bPullFail := FALSE;                 // 抽检失败预清零（独立记账）
_bAnyNg := FALSE;                    // 通道 NG 预清零
_bCfgBad := FALSE;                   // 组态非法预清零
nErrId := 16#0000_0000;              // 事件码缺省无事件
FOR _nK := 0 TO (nMaxCh - 1) DO
    abChannelOk[_nK] := FALSE;       // 通道结论缺省 FALSE（安全侧，段 3 单点置位）
    abPeakViolate[_nK] := FALSE;     // 峰值越窗缺省 FALSE
    abSlopeViolate[_nK] := FALSE;    // 斜率越窗缺省 FALSE
END_FOR

(* —— 段 2：组态域闸（覆盖全部参与判据换算的引脚，R151） —— *)
IF (nChannelCount <= 0) OR (nChannelCount > nMaxCh) THEN
    _bCfgBad := TRUE;                // 通道数越域（超 32 禁生成掩码，规格强制）
END_IF
IF (fPeakMaxC <= fPeakMinC) OR (fSlopeMaxCs <= fSlopeMinCs)
   OR (fHoldMaxMs <= fHoldMinMs) OR (fPullMinN <= 0.0) THEN
    _bCfgBad := TRUE;                // 判据窗倒置或拉力下限非法
END_IF
IF _bCfgBad THEN
    nErrId := 16#0006_02B4;          // 故障级：组态非法
    RETURN;                          // 不进入判据（出口维持安全缺省）
END_IF

(* —— 段 3：逐通道三判据（峰值窗 / 斜率窗 / 保温时长窗）+ SHL 显式位号聚合 —— *)
FOR _nK := 0 TO (nChannelCount - 1) DO
    _bFin := (afPeakC[_nK] = afPeakC[_nK]) AND (afSlopeCs[_nK] = afSlopeCs[_nK])
             AND (afHoldMs[_nK] = afHoldMs[_nK])
             AND (ABS(afPeakC[_nK]) < 1.0E6) AND (ABS(afSlopeCs[_nK]) < 1.0E6)
             AND (ABS(afHoldMs[_nK]) < 1.0E9);      // NaN 用 x<>x 自反，Inf 用幅值上限兜
    IF NOT _bFin THEN
        abChannelOk[_nK] := FALSE;      // 非有限通道按 NG 记（安全侧）
        abPeakViolate[_nK] := TRUE;     // 归入峰值越窗位段（头注释已声明）
        _uInfo := 16#0006_04B4;         // 信息级：非有限信号通道
    ELSE
        IF (afPeakC[_nK] < fPeakMinC) OR (afPeakC[_nK] > fPeakMaxC) THEN
            abPeakViolate[_nK] := TRUE; // 峰值越窗
        END_IF
        IF (afSlopeCs[_nK] < fSlopeMinCs) OR (afSlopeCs[_nK] > fSlopeMaxCs) THEN
            abSlopeViolate[_nK] := TRUE;    // 斜率越窗
        END_IF
        IF (afHoldMs[_nK] < fHoldMinMs) OR (afHoldMs[_nK] > fHoldMaxMs) THEN
            abPeakViolate[_nK] := TRUE;     // 保温时长越窗并入峰值位段（规格三判据聚合声明）
        END_IF
        abChannelOk[_nK] := (NOT abPeakViolate[_nK]) AND (NOT abSlopeViolate[_nK]);   // 通道结论
    END_IF
    IF NOT abChannelOk[_nK] THEN
        nNgChannelMask := nNgChannelMask OR SHL(DWORD(1), UINT(_nK));   // SHL 显式位号（禁魔法掩码）
        _bAnyNg := TRUE;                // 通道 NG 聚合（独立记账）
    END_IF
END_FOR
IF _bAnyNg THEN
    _uInfo := 16#0006_03B4;             // 信息级：存在曲线越窗通道
END_IF

(* —— 段 4：拉力抽检（仅抽中通道生效，独立记账不互相掩盖） —— *)
FOR _nK := 0 TO (nChannelCount - 1) DO
    IF abPullSampled[_nK] THEN
        IF (afPullN[_nK] <> afPullN[_nK]) OR (afPullN[_nK] < fPullMinN) THEN
            _bPullFail := TRUE;         // 抽检不合格（非有限按不合格记，安全侧）
        END_IF
    END_IF
END_FOR

(* —— 段 5：出口单点映射（名实同源；双判据独立记账，禁互相掩盖） —— *)
bLotReject := _bPullFail OR _bAnyNg;    // 整批判废：抽检失败或存在 NG 通道（任一成立）
IF _bPullFail THEN
    _uInfo := 16#0006_01B4;             // 信息级：抽检不合格整批判废
END_IF
IF _uInfo <> 16#0000_0000 THEN
    nErrId := _uInfo;                   // 信息码
END_IF

END_FUNCTION_BLOCK
